(* IEC 61131-3 sources: LASAL/Class/Varan_Base, 1 file *)

(* ---- Varan_Base.st ---- *)
#ifndef _T_VARANBASE_H
#define _T_VARANBASE_H

#define	VARAN_PLL_OFFSET		16#0140
#define VARAN_MULTIPLE_OFFSET	16#01AC

// version of serial number validation (16#10 = 1.0)
#define SERNO_VALIDATION_VERSION 16#10

#define IsTransparent_IS_AVAILABLE

// Defines for Mutex Generation
#define VARAN_STR_MUTEX_NAME_SEPERATOR ".."
#define VARAN_MUTEX_NAME_END_LENGTH 5
#define VARAN_MUTEX_NAME_MAX_LENGTH 32

#define VARAN_SPI_IDENT_LICENCENO_OFFSET    16#14
#define VARAN_SPI_IDENT_HARDWAREVER_OFFSET  16#18

#endif // _T_VARANBASE_H

#include "..\..\Class\HwControl\HwControl.h"
#include "..\..\Source\interfaces\lsl_st_hardwaretree.h"

(*!
<Class
	Name               = "Varan_Base"
	Revision           = "2.15"
	RealtimeTask       = "false"
	CyclicTask         = "false"
	BackgroundTask     = "false"
	Sigmatek           = "true"
	OSInterface        = "false"
	HighPriority       = "false"
	Automatic          = "false"
	UpdateMode         = "Prescan"
	IconPath           = ".\Class\Varan_Base\tool.ICO"
	SharedCommandTable = "true"
	Objectsize         = "(468,120)"
	Comment            = "baseclass of varan slave classes">
	<Channels>
		<Server Name="ConnectCounter" Visualized="true" Initialize="false" WriteProtected="true" Retentive="false" Comment="Connects of Module"/>
		<Server Name="DeviceAddress" Visualized="true" Initialize="false" WriteProtected="true" Retentive="false" Comment="device address of hardware module"/>
		<Server Name="DeviceID" Visualized="true" Initialize="false" WriteProtected="true" Retentive="false" Comment="This server shows the device ID of the hardware module."/>
		<Server Name="DiagControl" Visualized="true" Initialize="false" WriteProtected="false" Retentive="false" Comment="Server to control Diagnose Function of module&#13;&#10;&#13;&#10;Read from Server&#13;&#10;-2..wrong FPGA for Diagnose&#13;&#10;-1..wrong OS for Diagnose&#13;&#10;0..Diagnose Function is deaktivated, not available&#13;&#10;1..Diagnose Function activated (additionally you need #define VARAN_DIAGNOSE)&#13;&#10;&#13;&#10;Write to Server&#13;&#10;0..to deactivate Diagnose&#13;&#10;1..to activate Diagnose&#13;&#10;2..to reset Counter (ConnectCounter, FaultCounter, RXLost, TXLost)"/>
		<Server Name="FaultCounter" Visualized="true" Initialize="false" WriteProtected="true" Retentive="false" Comment="PackageCounter for RXLost and TXLost were invalid"/>
		<Server Name="Online" Visualized="true" Initialize="false" WriteProtected="true" Retentive="false" Comment="is class online or not"/>
		<Server Name="Release" Visualized="true" Initialize="false" WriteProtected="true" Retentive="false" Comment="FPGA - Version"/>
		<Server Name="RetryCounter" Visualized="true" Initialize="false" WriteProtected="false" Retentive="false" Comment="retry counter of varan module"/>
		<Server Name="RXLost" Visualized="true" Initialize="false" WriteProtected="true" Retentive="false" Comment="RX-Packages lost"/>
		<Server Name="SerialNo" Class="String" Visualized="true" Initialize="false" WriteProtected="true" Retentive="false" Comment="use this channel to access the string functions"/>
		<Server Name="State" Visualized="true" Initialize="false" WriteProtected="true" Retentive="false" Comment="This server shows the current status of the hardware class. For more information see: Varan hardware class status."/>
		<Server Name="TXLost" Visualized="true" Initialize="false" WriteProtected="true" Retentive="false" Comment="TX-Packages lost"/>
		<Server Name="ValidateSerNo" Visualized="true" Initialize="false" WriteProtected="false" Retentive="false" Comment="if the validation of the serial number is activated (SerNoValidation = 1)&#13;&#10;the serial number of the actual module can be validated by writing to this server&#13;&#10;&#13;&#10;this server shows also the state of validation:&#13;&#10;-2..validation not acivated&#13;&#10;-1..no module validated on this position&#13;&#10; 0..module is not the validated one&#13;&#10; 1..module is the validated one"/>
		<Server Name="VendorID" Visualized="true" Initialize="false" WriteProtected="true" Retentive="false" Comment="This server contains the vendor ID of the hardware module."/>
		<Client Name="Required" Required="true" Internal="false" Comment="0 = module is not required&#13;&#10;1 = module is required (CPU will crash if module is missing)"/>
		<Client Name="SerialNoStr" Required="true" Internal="true"/>
		<Client Name="SerNoBackup" Required="true" Internal="true"/>
		<Client Name="SerNoValidation" Required="false" Internal="false" Comment="0..serial number of varan client does not matter&#13;&#10;1..serial number of varan client has to be validated, to use the module&#13;&#10;&#13;&#10;validation is done via write(1) to the ValidateSerNo Server"/>
		<Client Name="TimeBase" Required="false" Internal="false" DefValue="0"/>
		<Client Name="TimeBaseOffset" Required="false" Internal="false" DefValue="0"/>
		<Client Name="To_MultiTask" Required="false" Internal="false" Comment="This client is automatically connected to a OS interface class."/>
		<Client Name="To_StdLib" Required="false" Internal="false" Comment="This client is automatically connected to a OS interface class."/>
		<Client Name="Transparent" Required="false" Internal="false" DefValue="0" Comment="If this Client is set to 1 the module is not used for building the VARAN-Tree"/>
		<Client Name="UserAction" Required="false" Internal="false" Comment="optional, connect to server to get Varan states via write method.&#13;&#10;possible input values:&#13;&#10; 0..connect&#13;&#10; 1..disconnect&#13;&#10; 2..required data object error&#13;&#10; 3..not required data object error&#13;&#10; 4..fatal error&#13;&#10; 5..time slice error&#13;&#10; 6..watchdog error&#13;&#10; 7..client irq&#13;&#10; 8..device enable&#13;&#10; 9..device disable&#13;&#10;10..irq task interrupt&#13;&#10;11..reactivation of node which was deactivated by software before&#13;&#10;12..irq for direct access alternating buffer (VMC module)&#13;&#10;13..dias error&#13;&#10;14..cdias error (cdias module required behind a CIV)&#13;&#10;&#13;&#10;&#13;&#10;Possible return values:&#13;&#10;0......ok&#13;&#10;&lt;&gt; 0...Generate VaranError&#13;&#10;"/>
		<Client Name="VaranIn" Required="true" Internal="false" Comment="This class must be connected to a VARAN port or a VaranOut_[x] server."/>
	</Channels>
	<Dependencies>
		<Files>
			<File Path=".\Class\VaranManager_Base\VaranManager_Base.h" Include="false"/>
			<File Path=".\Source\interfaces\lsl_st_pci.h" Include="false"/>
			<File Path=".\Class\HwControl\HwControl.h" Include="true"/>
			<File Path=".\Source\interfaces\lsl_st_hardwaretree.h" Include="true"/>
		</Files>
	</Dependencies>
	<RevDoku>
		<Owner Company="Sigmatek" Author="renste"/>
		<Dokumentation Revision="2.15" Date="16.03.2018" Author="EisMic" Company="Sigmatek" Description="Added support for 2nd VaranManager."/>
		<Dokumentation Revision="2.14" Date="06.03.2018" Author="EisMic" Company="Sigmatek" Description="Attached header files no longer point to the installation directory of LASAL but instead now point to the the source/interfaces folder."/>
		<Dokumentation Revision="2.13" Date="10.01.2018" Author="LanSte" Company="Sigmatek" Description="Added Support for default PostInit phase."/>
		<Dokumentation Revision="2.12" Date="23.01.2018" Author="RamAnd" Company="Sigmatek" Description="Log messages have been standardized for easier maintenance, easier use in any class and to allow spam filtering. Code for the logging functions is now only located in HwControl."/>
		<Dokumentation Revision="2.11" Date="28.08.2017" Author="RamAnd" Company="Sigmatek" Description="The NewInst to get hardware diagnosis information doesn&apos;t set the returncode to SPI_ACCESS_FAILED if an optional entry of the type label is not available."/>
		<Dokumentation Revision="2.10" Date="29.11.2016" Author="PieSte" Company="Sigmatek" Description="Changed &quot;Online&quot; server behavior to set online first if cyclic data is valid."/>
		<Dokumentation Revision="2.9" Date="10.05.2016" Author="RamAnd" Company="Sigmatek" Description="Suppressed warning that would occur with target ARM on compiler version 30 or higher."/>
		<Dokumentation Revision="2.8" Date="17.02.2016" Author="EisMic" Company="Sigmatek" Description="Prescalersettings were not set correctly when Payload is active."/>
		<Dokumentation Revision="2.7" Date="28.08.2015" Author="PieSte" Company="Sigmatek" Description="Added support for up to 6 sync outs (e.g. CTMS031) in methode EnableSyncOut()."/>
		<Dokumentation Revision="2.6" Date="17.03.2015" Author="RamAnd" Company="Sigmatek" Description="Added support for Varan Mux."/>
		<Dokumentation Revision="2.5" Date="24.03.2015" Author="EisMic" Company="Sigmatek" Description="Check pointer p_NodeInfo for validity in method GetRetryTimeout due to access exception error if method Varan_HWDisconnect is called and no hardware was available."/>
		<Dokumentation Revision="2.4" Date="28.08.2014" Author="EisMic" Company="Sigmatek" Description="Don&apos;t set states in GetHWInfoData. CMD_Get_Hardware_Diagnosis: Don&apos;t do a return when one spi access failed, try the other IDs too."/>
		<Dokumentation Revision="2.3" Date="24.06.2014" Author="LanSte" Company="Sigmatek" Description="Added support for reading hardware diagnosis."/>
		<Dokumentation Revision="2.2" Date="05.05.2014" Author="LanSte" Company="Sigmatek" Description="Minimized the interface request via CILGET by useing private pointers to reduce time in init."/>
		<Dokumentation Revision="2.1" Date="14.04.2014" Author="RamAnd" Company="Sigmatek" Description="Added new Interface Varan_HwSubBusReady which is called by OS as soon as it has finished enumerating the connected devices on available subbusses."/>
		<Dokumentation Revision="2.0" Date="04.12.2013" Author="RamAnd&#13;&#10;FucHer&#13;&#10;LanSte" Company="Sigmatek" Description="Removed domain support&#13;&#10;Changed AWL code to Structured Text.&#13;&#10;Added Payload Support&#13;&#10;Added include for PCI accesses, which is necessary to find out if the Varan Manager supports LongDOs."/>
		<Dokumentation Revision="1.90" Date="30.08.2013" Author="RamAnd" Company="Sigmatek" Description="The class could have change the state to _DisableError after the disconnect from VARAN, even if there was no further problem."/>
		<Dokumentation Revision="1.80" Date="01.08.2013" Author="LanSte" Company="Sigmatek" Description="Added Support for changeable Payload DO&apos;s"/>
		<Dokumentation Revision="1.70" Date="18.07.2013" Author="LanSte&#13;&#10;ZoePat" Company="Sigmatek" Description="Added Payload Support&#13;&#10;Check if manager is on at function GetNodeInfo() to get different states for connected and disconnected modules if manager is turned off (e.g.: in case of required error that was handled by client UserAction)"/>
		<Dokumentation Revision="1.60" Date="07.03.2013" Author="RamAnd" Company="Sigmatek" Description="Improved comment of client UserAction (added new reasons)"/>
		<Dokumentation Revision="1.50" Date="05.11.2012" Author="RamAnd&#13;&#10;RamAnd" Company="Sigmatek" Description="Corrected time measurement for internal tests.&#13;&#10;Removed resetting of the FPGA retry counter in method ResetDataObject which could result in a wrong behavior of the RetryCounter server."/>
		<Dokumentation Revision="1.40" Date="18.09.2012" Author="RamAnd" Company="Sigmatek" Description="New State &quot;_NoCalibDataFound&quot; if a pointer to calibration data is fetched and there are no calibration data on the client."/>
		<Dokumentation Revision="1.39" Date="18.07.2012" Author="ObeChr" Company="Sigmatek" Description="Implemented time measurement for internal tests in methods UpdateRt, UpdateRtPostScan and UpdateCy&#13;&#10;Reduction of PCI Accesses in Methode GetRetryTimeout()"/>
		<Dokumentation Revision="1.38" Date="09.12.2011" Author="RamAnd" Company="Sigmatek" Description="The actual domain number is now added to the hardware path."/>
		<Dokumentation Revision="1.37" Date="19.09.2011" Author="RamAnd" Company="Sigmatek" Description="The client UserAction can now also be used to prevent a required error, if the write-method of the connected Server returns 0."/>
		<Dokumentation Revision="1.36" Date="13.07.2011" Author="RamAnd" Company="Sigmatek" Description="Added a dependency to class Hub_Base_Root, otherwise crashes can happen if only single VARAN-classes have been updated."/>
		<Dokumentation Revision="1.35" Date="14.04.2011" Author="BleErn" Company="Sigmatek" Description="Set complex object &quot;SerialNoStr&quot; to visualized"/>
		<Dokumentation Revision="1.34" Date="02.03.2011" Author="RamAnd" Company="Sigmatek" Description="Added new input parameter to method SetMultipleDataPointers to handle more than 1 multiple read write commands per VARAN client."/>
		<Dokumentation Revision="1.33" Date="04.01.2011" Author="BleErn" Company="Sigmatek" Description="Added Client Transparent that allows to disable a VARAN-HW-Class"/>
		<Dokumentation Revision="1.32" Date="17.01.2011" Author="RamAnd" Company="Sigmatek" Description="A required error on the first connect of the device can now be detected via the UserAction client"/>
		<Dokumentation Revision="1.31" Date="11.01.2011" Author="RamAnd" Company="Sigmatek" Description="Error fixed that Diagnostic functions stopped working after the first fault occured."/>
		<Dokumentation Revision="1.30" Date="14.12.2010" Author="RamAnd" Company="Sigmatek" Description="Set all servers to visualized, so that they can be used in visualisation"/>
		<Dokumentation Revision="1.29" Date="02.09.2010" Author="BleErn" Company="Sigmatek" Description="Server SerNoValidation was always set to 0 on disconnect of module"/>
		<Dokumentation Revision="1.28" Date="02.08.2010" Author="RamAnd" Company="Sigmatek" Description="Reworked serial number validation, because of problems with non-Sigmatek devices. Now the serial number is saved as a string instead of a number."/>
		<Dokumentation Revision="1.27" Date="22.07.2010" Author="WocPet / RamAnd" Company="Sigmatek" Description="Added functionality to forward a required error.&#13;&#10;Removed client UseRtPostScan (not needed, since it PostScan is always used)"/>
		<Dokumentation Revision="1.26" Date="06.04.2010" Author="RamAnd" Company="Sigmatek" Description="Added method &quot;FlexInit&quot; to initialize class if the position on VARAN has changed (FlexHub functionality)"/>
		<Dokumentation Revision="1.25" Date="10.03.2010" Author="RamAnd" Company="Sigmatek" Description="Added serial number validation and method CheckDeviceID for easier overloading"/>
		<Dokumentation Revision="1.24" Date="04.03.2010" Author="BleErn" Company="Sigmatek" Description="RtPostScan could be disabled at every CIV (took no notice of define!)"/>
		<Dokumentation Revision="1.23" Date="23.02.2010" Author="BleErn" Company="Sigmatek" Description="Changes in handling of VaranRtPostScan"/>
		<Dokumentation Revision="1.22" Date="17.05.2010" Author="RamAnd" Company="Sigmatek" Description="Changed defines to avoid compiler warning &quot;Identical Redefinition&quot;"/>
		<Dokumentation Revision="1.21" Date="09.10.2009" Author="ObeChr" Company="Sigmatek" Description="Added functions for VaranDiagnose"/>
		<Dokumentation Revision="1.20" Date="02.09.2009" Author="RamAnd" Company="Sigmatek" Description="Added functions for safety and hardwaretree."/>
		<Dokumentation Revision="1.19" Date="05.08.2009" Author="ObeChr" Company="Sigmatek" Description="When Client is required and no VaranInterface is available, VaranManager set application into reset"/>
		<Dokumentation Revision="1.18" Date="20.07.2009" Author="ObeChr" Company="Sigmatek" Description="Added function to set run state of do depending on required"/>
		<Dokumentation Revision="1.17" Date="16.07.2009" Author="ObeChr" Company="Sigmatek" Description="Added funktion to use VaranRtPostScan"/>
		<Dokumentation Revision="1.16" Date="18.06.2009" Author="EbnAnt" Company="Sigmatek" Description="Set Varan_CallBack() to virtual"/>
		<Dokumentation Revision="1.15" Date="16.04.2009" Author="RamAnd" Company="Sigmatek" Description="Added new method GetDocumentation to fetch pdf documentation of client.&#13;&#10;Added new Server SerialNo, to display the serial no of varan clients."/>
		<Dokumentation Revision="1.14" Date="01.12.2008" Author="RamAnd" Company="Sigmatek" Description="added new input variable b_use_divider_sync to function EnableSyncOut.&#13;&#10;Corrected SetNewPllData to new address mapping.&#13;&#10;improved client comments"/>
		<Dokumentation Revision="1.13" Date="03.09.2008" Author="renste" Company="Sigmatek" Description="add function for new pll"/>
	</RevDoku>
	<Network Name="Varan_Base">
		<!-- List of Components in this network -->
		<Components>
			<Object
				Name       = "SerialNoStr"
				Class      = "String"
				Position   = "(180,480)"
				Visualized = "true">
				<Channels>
					<Server Name="Data"/>
					<Client Name="SingleRealloc" Value="1"/>
				</Channels>
			</Object>
			<Object
				Name       = "SerNoBackup"
				Class      = "RamFile"
				Position   = "(180,630)"
				Visualized = "true">
				<Channels>
					<Server Name="FileNameHex"/>
					<Server Name="m_udLength"/>
					<Server Name="SizeError"/>
					<Client Name="Alarm"/>
					<Client Name="MultiTask"/>
					<Client Name="Setup" Value="2#1101"/>
				</Channels>
			</Object>
		</Components>
		<Comments>
		</Comments>
		<!-- List of Connections in this network -->
		<Connections>
			<Connection Source="this.SerialNoStr" Destination="SerialNoStr.Data"/>
			<Connection Source="this.SerialNo" Destination="SerialNoStr.Data" Vertices="(818,570),(496,570),"/>
			<Connection Source="this.SerNoBackup" Destination="SerNoBackup.m_udLength"/>
		</Connections>
		<!-- Headerfiles -->
		<Options>
		</Options>
	</Network>
</Class>
*)
Varan_Base : CLASS
	TYPE
	  t_CallBack : STRUCT
	    ud_Counter : UDINT;
	    ud_ConnectCnt : UDINT;
	    ud_DisconnectCnt : UDINT;
	    ud_InterruptCnt : UDINT;
	    ud_SubBusReadyCnt : UDINT;
	    p_InterruptHandleDO : ^LSL_VARANFRAME;  //! <Type Comment="Warning:&#13;&#10;If the Interface &quot;IMULTIVARANMANAGER&quot; is used (b_PayloadSupport = true) this pointer those not point to the DO in the DPRAM!&#13;&#10;In this case this pointer holds the handle to the DO.&#13;&#10;" Name="t_CallBack.p_InterruptHandleDO"/>
	    ud_LastReason : UDINT;
	  END_STRUCT;
	  t_CycleWork :
	  (
	    _CycleInitIdle,
	    _CycleStartAsyDO,
	    _CycleStartIsoDO,
	    _CycleWaitforValidData,
	    _CyclePreOperational,
	    _CycleOperational
	  )$UDINT;
	  t_PllDataRead : STRUCT
	    us_State : BSINT
	    [
	      1 Pll_Locked,
	      2 Pll_Unlocked,
	      3 SyncOutputAvailable0,
	      4 SyncOutputAvailable1,
	      5 SyncOutputAvailable2,
	      6 IRQWatchdogEnable,
	      7 Pll_Enable,
	      8 PeriodeOverwriteAllowed,
	    ];
	  END_STRUCT;
	  t_PllDO : STRUCT
	    p_Handle : ^LSL_VARANFRAME;
	    p_DOSettings : ^t_VaranDOSettingsRd;
	    p_DataRead : ^t_PllDataRead;
	  END_STRUCT;
#pragma pack(push, 1)
	  t_PllSyncOut : STRUCT
	    sd_Offset : DINT;
	    us_PeriodMultiplier : USINT;
	    us_FrameCountTreshold : USINT;
	    us_Reserved1 : USINT;
	    us_ControlStatus : BSINT
	    [
	      1 SyncOutEnable,
	      2 FrameCountEnable,
	      3 SystemSync,  //! <Type Comment="0..divider sync&#13;&#10;1..system sync" Name="t_PllSyncOut.us_ControlStatus.SystemSync"/>
	    ];
	  END_STRUCT;
#pragma pack(pop)
	  t_RootDependency : ^Hub_Base_Root;
#pragma pack(push, 1)
	  t_SerNoValidateHeader : STRUCT
	    Version : HSINT;  //! <Type Comment="X.Y starting with 1.0 as first valid version&#13;&#10;&#13;&#10;X = Major&#13;&#10;Y = Minor" Name="t_SerNoValidateHeader.Version"/>
	    ZeroByte : USINT;
	    StringLength : UDINT;
	  END_STRUCT;
#pragma pack(pop)
	  t_SPI_CalibHeader : STRUCT
	    ud_Checksum : UDINT;
	    ud_ListVersion : UDINT;
	    ud_ListLength : UDINT;
	  END_STRUCT;
	  t_TempDataRead : STRUCT
	    si_Periode : INT;
	    ui_Prescaler : UINT;
	    ui_HiTimeRegister : UINT;
	  END_STRUCT;
	  t_TransparentInfo : BSINT
	  [
	    1 DeviceIsTransparent,
	    2 ClientTransparentRead,
	  ];
	END_TYPE
  //Servers:
	State 	: SvrChCmd_t_e_VaranErrors;
	Online 	: SvrCh_DINT;
	Release 	: SvrCh_HDINT;
	DeviceAddress 	: SvrCh_HDINT;
	VendorID 	: SvrCh_UDINT;
	DeviceID 	: SvrCh_UDINT;
	SerialNo 	: SvrChCmd_UDINT;
	RetryCounter 	: SvrCh_UDINT;
	ValidateSerNo 	: SvrCh_DINT;
	DiagControl 	: SvrCh_DINT;
	ConnectCounter 	: SvrCh_UDINT;
	FaultCounter 	: SvrCh_UDINT;
	RXLost 	: SvrCh_UDINT;
	TXLost 	: SvrCh_UDINT;
  //Clients:
	VaranIn 	: CltChCmd_Hub_Base;
	Required 	: CltCh_DINT;
	UserAction 	: CltCh_DINT;
	SerNoValidation 	: CltCh_DINT;
	Transparent 	: CltCh_DINT;
	To_StdLib 	: CltChCmd__StdLib;
	To_MultiTask 	: CltChCmd__MultiTask;
	TimeBase 	: CltCh_UDINT;
	TimeBaseOffset 	: CltCh_UDINT;
	SerialNoStr 	: CltChCmd_String;
	SerNoBackup 	: CltChCmd_RamFile;
  //Variables:
		ud_VaranManagerNr 	: UDINT;
		pVaran 	: ^LSL_VARAN;			//! <Variable Comment="Pointer for the Varan interface" Name="pVaran"/>
		pMultiVaran 	: ^LSL_MULTI_VARAN;			//! <Variable Comment="Pointer for the MultiVaran/payload support interface" Name="pMultiVaran"/>
		mt_api 	: ^LSL_MT_TYPE;
		p_VaranPosition 	: ^USINT;
		p_NodeInfo 	: ^LSL_VARANNODEINFO;
		s_NodeInfo 	: LSL_VARANNODEINFO;
		ud_HandleModule 	: UDINT;
		ud_DeviceDelayTime 	: UDINT;
		s_CallBackSettings 	: t_CallBack;			//! <Variable Comment="settings of user callback function" Name="s_CallBackSettings"/>
		e_RequiredFaultState 	: t_e_VaranErrors;
		b_DisableDevice 	: BOOL;
		ud_DisableTime 	: UDINT;
		us_MulticastFilter 	: USINT;
		us_MultipleSequence 	: USINT;
		s_TimeRt 	: t_TimeMeasurementVaran;
		s_TimeRtPostScan 	: t_TimeMeasurementVaran;
		s_TimeCy 	: t_TimeMeasurementVaran;
		b_CyTask 	: BOOL;
		p_ObjectPath 	: ^USINT;
		s_Diagnose 	: t_s_VaranDiagnose;
		szSerNoStr : ARRAY [0..SERNO_STRING_SIZE-1] OF CHAR;

		b_ValidationInProgress 	: BOOL;
		SerNoHeader 	: t_SerNoValidateHeader;
		TransparentInfo 	: t_TransparentInfo;
		ud_ResponseTimeMax 	: UDINT;
		b_PayloadSupport 	: BOOL;			//! <Variable Comment="TRUE When Payload DOs are supporded by the OS Interface." Name="b_PayloadSupport"/>
		b_DMAactive 	: BOOL;			//! <Variable Comment="TRUE When Payload DOs are supporded by the OS Interface and the FPGA has an DMA Controller." Name="b_DMAactive"/>
		ud_OffestSPI 	: UDINT;
		bOnline 	: BOOL;
		eCycleWork 	: t_CycleWork;
		uiBasePostInitHandle 	: UINT;
		bPostInitNeeded 	: BOOL;
		_ParaBaseCy 	: CmdStruct;
		_ResultBaseCy 	: results;
  //Functions:
				//! <Function Comment="-------------------------------------------------------------------------------------------------&#13;&#10;[#ENGLISH]&#13;&#10;=================================================================================================&#13;&#10;Construct of Base class to set class not initialized&#13;&#10;=================================================================================================&#13;&#10;[server] State  :W  :State of class&#13;&#10;" Name="Varan_Base"/>
	FUNCTION Varan_Base
		VAR_OUTPUT
			ret_code 	: ConfStates;
		END_VAR;
				//! <Function Comment="Init for Varan Client" Name="Init"/>
	FUNCTION VIRTUAL GLOBAL Init;
				//! <Function Comment="Cy - Funktion of Varan class ( called bei VaranMaster )" Name="UpdateCy"/>
	FUNCTION VIRTUAL GLOBAL UpdateCy;
				//! <Function Comment="Rt - Funktion of Varan class ( called bei VaranMaster )" Name="UpdateRt"/>
	FUNCTION VIRTUAL GLOBAL UpdateRt;
				//! <Function Comment="Function is called by VaranRtPostScan if used" Name="UpdateRtPostScan"/>
	FUNCTION VIRTUAL GLOBAL UpdateRtPostScan;
				//! <Function Comment="get PDF-File from client, if it is available" Name="GetDocumentation"/>
	FUNCTION VIRTUAL GLOBAL GetDocumentation
		VAR_INPUT
			p_dpne 	: ^CHAR;			//! <Variable Comment="pass string of Drive/Path/Name/Extension (e.g. &quot;C:\mydoc.pdf&quot;)" Name="GetDocumentation.p_dpne"/>
		END_VAR
		VAR_OUTPUT
			sd_retval 	: DINT;			//! <Variable Comment=" 0..success&#13;&#10;-1..invalid parameters&#13;&#10;-2..failed to open file&#13;&#10;-3..os version must be 01.02.018 or higher&#13;&#10;-4..no documentation available on this client&#13;&#10;-5..failed to allocate memory for the file content&#13;&#10;-6..error in reading documentation from client&#13;&#10;-7..writing to file failed" Name="GetDocumentation.sd_retval"/>
		END_VAR;
				//! <Function Comment="Function returns pointer to node string of class" Name="GetPointer2NodeString"/>
	FUNCTION VIRTUAL GLOBAL GetPointer2NodeString
		VAR_OUTPUT
			p_us_node 	: ^USINT;			//! <Variable Comment="pointer to node string" Name="GetPointer2NodeString.p_us_node"/>
		END_VAR;
				//! <Function Comment="Function is called if a varan module is connected&#13;&#10;" Name="Varan_HwConnect"/>
	FUNCTION VIRTUAL GLOBAL Varan_HwConnect
		VAR_INPUT
			ud_data 	: UDINT;			//! <Variable Comment="data of callback function" Name="Varan_HwConnect.ud_data"/>
		END_VAR
		VAR_OUTPUT
			sd_retval 	: DINT;			//! <Variable Comment="return value of OS" Name="Varan_HwConnect.sd_retval"/>
		END_VAR;

	FUNCTION Diagnose;
				//! <Function Comment="[#ENGLISH]&#13;&#10;=================================================================================================&#13;&#10;Function to set Pll settings of hardware module&#13;&#10;=================================================================================================&#13;&#10;[server] State    :W  :state of class&#13;&#10;[members] ud_DeviceDelayTime :W  :delay time of varan client for Pll&#13;&#10;   p_NodeInfo   :W  :pointer to varan client informations&#13;&#10;[locals] ud_data    :W/R :data for direct access&#13;&#10;" Name="SetPllData"/>
	FUNCTION SetPllData
		VAR_INPUT
			ud_delay_time 	: UDINT := 0;
		END_VAR
		VAR_OUTPUT
			sd_retval 	: DINT;
		END_VAR;
				//! <Function Comment="[#ENGLISH]&#13;&#10;=================================================================================================&#13;&#10;Function to get device address, Vendor ID and Device ID of varan module&#13;&#10;=================================================================================================&#13;&#10;[server] State   :W  :state of class&#13;&#10;   Release   :W  :FPGA - Version of varan client&#13;&#10;   DeviceAddress :W  :Device Address of client (from os)&#13;&#10;   VendorID  :W  :Vendor ID of varan client&#13;&#10;   DeviceID  :W  :Device ID of varan client&#13;&#10;[members] p_VaranPosition  :R  :node string of varan module&#13;&#10;   p_NodeInfo   :W  :pointer to varan client informations&#13;&#10;[locals] us_pll_time   :W/R :pll time from VaranMaster&#13;&#10;" Name="GetNodeInfo"/>
	FUNCTION GetNodeInfo
		VAR_OUTPUT
			sd_retval 	: DINT;
		END_VAR;
				//! <Function Comment="[#ENGLISH]&#13;&#10;=================================================================================================&#13;&#10;Callback Function is called from VaranManager&#13;&#10;=================================================================================================&#13;&#10;[server] Release   :W  :FPGA - Version of varan client&#13;&#10;   DeviceAddress :W  :Device Address of client (from os)&#13;&#10;   VendorID  :W  :Vendor ID of varan client&#13;&#10;   DeviceID  :W  :Device ID of varan client&#13;&#10;   State   :W  :state of class&#13;&#10;[client] Required  :R  :is class required for varan or not&#13;&#10;   UserAction  :R  :client for user actions&#13;&#10;[members] s_CallBackSettings  :W  :structure for settings of callback function&#13;&#10;   ud_DeviceDelayTime  :W  :delay time of varan client for Pll&#13;&#10;   e_RequiredFaultState :W  :Fault state of class in _RequiredError State&#13;&#10;" Name="Varan_CallBack"/>
	FUNCTION VIRTUAL Varan_CallBack
		VAR_INPUT
			ud_reason 	: UDINT;			//! <Variable Comment="reason of callback" Name="Varan_CallBack.ud_reason"/>
			ud_data 	: UDINT;
		END_VAR
		VAR_OUTPUT
			sd_retval (EAX) 	: DINT;
		END_VAR;
				//! <Function Comment="Function is called if a varan interrupt occures" Name="Varan_HwInterrupt"/>
	FUNCTION VIRTUAL GLOBAL Varan_HwInterrupt
		VAR_INPUT
			ud_reason 	: UDINT;
			ud_data 	: ^t_CallBackInterrupt;
		END_VAR
		VAR_OUTPUT
			sd_retval 	: DINT;
		END_VAR;
				//! <Function Comment="Function is called if a varan module is disconnected&#13;&#10;" Name="Varan_HwDisconnect"/>
	FUNCTION VIRTUAL GLOBAL Varan_HwDisconnect
		VAR_INPUT
			ud_data 	: UDINT;
		END_VAR
		VAR_OUTPUT
			sd_retval 	: DINT;
		END_VAR;

	FUNCTION VIRTUAL GLOBAL Varan_HwSubBusReady
		VAR_INPUT
			ud_data 	: UDINT;
		END_VAR
		VAR_OUTPUT
			sd_retval 	: DINT;
		END_VAR;
				//! <Function Comment="Function to reset settings of a data object" Name="ResetDataObject"/>
	FUNCTION VIRTUAL GLOBAL ResetDataObject
		VAR_INPUT
			p_handleDO 	: ^LSL_VARANFRAME;
			us_state 	: USINT;			//! <Variable Comment="state of DO (cont run, singl run, stop )" Name="ResetDataObject.us_state"/>
			ud_bytes 	: UDINT;			//! <Variable Comment="number of bytes" Name="ResetDataObject.ud_bytes"/>
		END_VAR;
				//! <Function Comment="=================================================================================================&#13;&#10;---------------------- Additional functions------------------------------------------------------&#13;&#10;=================================================================================================&#13;&#10;[#ENGLISH]&#13;&#10;=================================================================================================&#13;&#10;Function to Start time measurement&#13;&#10;=================================================================================================&#13;&#10;" Name="StartTimeMeasurement"/>
	FUNCTION StartTimeMeasurement
		VAR_INPUT
			usMode (EAX) 	: DINT;
		END_VAR;
				//! <Function Comment="[#ENGLISH]&#13;&#10;=================================================================================================&#13;&#10;Function to Stop time measurement&#13;&#10;=================================================================================================&#13;&#10;" Name="StopTimeMeasurement"/>
	FUNCTION StopTimeMeasurement
		VAR_INPUT
			usMode (EAX) 	: DINT;
		END_VAR;
				//! <Function Comment="Function to set a sync out" Name="GetDeviceAddress"/>
	FUNCTION VIRTUAL GLOBAL GetDeviceAddress
		VAR_OUTPUT
			ud_device_address 	: UDINT;			//! <Variable Comment="Device address of client" Name="GetDeviceAddress.ud_device_address"/>
		END_VAR;
				//! <Function Comment="[#ENGLISH]&#13;&#10;=================================================================================================&#13;&#10;Function to set a sync out&#13;&#10;=================================================================================================&#13;&#10;[server] State    :W  :state of class&#13;&#10;[locals] ud_offset    :W/R :address offset in pll&#13;&#10;   p_pll_output_data  :W/R :settings for pll sync output&#13;&#10;" Name="EnableSyncOut"/>
	FUNCTION EnableSyncOut
		VAR_INPUT
			us_sync_nr 	: USINT;			//! <Variable Comment="enable sync0-4 allowed" Name="EnableSyncOut.us_sync_nr"/>
			sd_offset 	: DINT;			//! <Variable Comment="Offset in 10ns time" Name="EnableSyncOut.sd_offset"/>
			us_period_multiplier 	: USINT;			//! <Variable Comment="periode multiplier" Name="EnableSyncOut.us_period_multiplier"/>
			us_frame_count_treshold 	: USINT;			//! <Variable Comment=" Frame Count Treshold" Name="EnableSyncOut.us_frame_count_treshold"/>
			us_enable_frame_count 	: USINT;			//! <Variable Comment=" enable frame count" Name="EnableSyncOut.us_enable_frame_count"/>
			b_use_divider_sync 	: BOOL := FALSE;
		END_VAR
		VAR_OUTPUT
			sd_retval 	: DINT;
		END_VAR;
				//! <Function Comment="Function to get pointer to node information" Name="GetPointer2NodeInfo"/>
	FUNCTION VIRTUAL GLOBAL GetPointer2NodeInfo
		VAR_OUTPUT
			p_node_info 	: ^LSL_VARANNODEINFO;			//! <Variable Comment="Pointer to Node information" Name="GetPointer2NodeInfo.p_node_info"/>
		END_VAR;
				//! <Function Comment="Function to set state of class" Name="SetState"/>
	FUNCTION VIRTUAL GLOBAL SetState
		VAR_INPUT
			sd_error 	: t_e_VaranErrors;			//! <Variable Comment="type of error" Name="SetState.sd_error"/>
		END_VAR;
				//! <Function Comment="Function to disable device" Name="DisableDevice"/>
	FUNCTION VIRTUAL GLOBAL DisableDevice
		VAR_OUTPUT
			sd_retval 	: DINT;
		END_VAR;
				//! <Function Comment="Function to enable device" Name="EnableDevice"/>
	FUNCTION VIRTUAL GLOBAL EnableDevice
		VAR_OUTPUT
			sd_retval 	: DINT;
		END_VAR;
				//! <Function Comment="Function to set all Data Objects off" Name="SetDOsOff"/>
	FUNCTION VIRTUAL GLOBAL SetDOsOff;
				//! <Function Comment="Function to look if class is disabled" Name="IsDeviceDisabled"/>
	FUNCTION VIRTUAL GLOBAL IsDeviceDisabled
		VAR_OUTPUT
			b_disabled 	: BOOL;			//! <Variable Comment="TRUE -&gt; Device is disabled" Name="IsDeviceDisabled.b_disabled"/>
		END_VAR;
				//! <Function Comment="Function to set multiple memory read/write options" Name="SetMultipleSettings"/>
	FUNCTION VIRTUAL GLOBAL SetMultipleSettings
		VAR_INPUT
			us_filter 	: USINT;			//! <Variable Comment="filter of multicast write" Name="SetMultipleSettings.us_filter"/>
			us_sequence 	: USINT;			//! <Variable Comment="sequence number of device" Name="SetMultipleSettings.us_sequence"/>
		END_VAR
		VAR_OUTPUT
			sd_retval 	: DINT;
		END_VAR;
				//! <Function Comment="Function must be overwrite" Name="SetMultipleDataPointers"/>
	FUNCTION VIRTUAL GLOBAL SetMultipleDataPointers
		VAR_INPUT
			p_handle 	: ^LSL_VARANFRAME;			//! <Variable Comment="pointer to data object header" Name="SetMultipleDataPointers.p_handle"/>
			p_data_read 	: ^UDINT;			//! <Variable Comment="pointer to read data" Name="SetMultipleDataPointers.p_data_read"/>
			p_data_write 	: ^UDINT;			//! <Variable Comment="pointer to data write" Name="SetMultipleDataPointers.p_data_write"/>
			DOIndex 	: UDINT;
		END_VAR
		VAR_OUTPUT
			sd_retval 	: DINT;
		END_VAR;
				//! <Function Comment="[#ENGLISH]&#13;&#10;=================================================================================================&#13;&#10;Function to get pointer to calib data&#13;&#10;=================================================================================================&#13;&#10;" Name="GetCalibDataPointer"/>
	FUNCTION GetCalibDataPointer
		VAR_INPUT
			p_offset 	: ^UDINT;			//! <Variable Comment="pointer to variable to write offset" Name="GetCalibDataPointer.p_offset"/>
		END_VAR
		VAR_OUTPUT
			sd_retval 	: DINT;
		END_VAR;
				//! <Function Comment="[#ENGLISH]&#13;&#10;=================================================================================================&#13;&#10;Function to get pointer to calib data&#13;&#10;=================================================================================================&#13;&#10;" Name="ReadSPIData"/>
	FUNCTION ReadSPIData
		VAR_INPUT
			ud_offset 	: UDINT;			//! <Variable Comment="offset in SPI - Flash" Name="ReadSPIData.ud_offset"/>
			ud_length 	: UDINT;			//! <Variable Comment="length of data" Name="ReadSPIData.ud_length"/>
			p_data 	: ^USINT;			//! <Variable Comment="pointer to allocated data space" Name="ReadSPIData.p_data"/>
		END_VAR
		VAR_OUTPUT
			sd_retval 	: DINT;
		END_VAR;
				//! <Function Comment="Function to update module retry counter" Name="UpdateRetryCounter"/>
	FUNCTION VIRTUAL GLOBAL UpdateRetryCounter;
				//! <Function Comment="Function to get varan time" Name="GetVaranTime"/>
	FUNCTION VIRTUAL GLOBAL GetVaranTime
		VAR_INPUT
			p_ud_IsoStartPoint 	: ^UDINT := NIL;
		END_VAR
		VAR_OUTPUT
			ud_varan_time 	: UDINT;			//! <Variable Comment="varan time" Name="GetVaranTime.ud_varan_time"/>
		END_VAR;
				//! <Function Comment="Function to get retry timeout for a number of bytes" Name="GetRetryTimeout"/>
	FUNCTION VIRTUAL GLOBAL GetRetryTimeout
		VAR_INPUT
			ud_bytes 	: UDINT;
		END_VAR
		VAR_OUTPUT
			ud_timeout 	: UDINT;			//! <Variable Comment="retry timout time" Name="GetRetryTimeout.ud_timeout"/>
		END_VAR;
				//! <Function Comment="[#ENGLISH]&#13;&#10;=================================================================================================&#13;&#10;Function to disable Device in Rt (because VARAN_iSetNodeEnableStatus must not called in Realtime)&#13;&#10;=================================================================================================&#13;&#10;" Name="DisableDeviceRt"/>
	FUNCTION DisableDeviceRt
		VAR_OUTPUT
			sd_retval 	: DINT;
		END_VAR;

	FUNCTION SetNewPllData
		VAR_INPUT
			ud_delay_time 	: UDINT := 0;
			us_divider 	: USINT := 0;
		END_VAR
		VAR_OUTPUT
			sd_retval 	: DINT;
		END_VAR;
				//! <Function Comment="Function to set state depending on required" Name="SetRunStatus"/>
	FUNCTION GLOBAL SetRunStatus
		VAR_INPUT
			state 	: USINT;
		END_VAR
		VAR_OUTPUT
			us_retval 	: USINT;
		END_VAR;

	FUNCTION VIRTUAL GLOBAL GetPointer2ObjectPath
		VAR_OUTPUT
			p_us_ObjectPath 	: ^USINT;
		END_VAR;

	FUNCTION VIRTUAL GLOBAL SetObjectThisp
		VAR_INPUT
			p_us_ObjectPath 	: ^USINT;
			ud_thisp 	: UDINT;
		END_VAR
		VAR_OUTPUT
			sd_retval 	: DINT;
		END_VAR;

	FUNCTION VIRTUAL GLOBAL GetObjectThisp
		VAR_INPUT
			p_us_ObjectPath 	: ^USINT;
		END_VAR
		VAR_OUTPUT
			ud_Thisp 	: UDINT;
		END_VAR;

	FUNCTION SerNoValidationTask;

	FUNCTION GetHWInfoData
		VAR_INPUT
			p_offset 	: ^UDINT;
			ud_id 	: UDINT;
		END_VAR
		VAR_OUTPUT
			sd_retval 	: DINT;
		END_VAR;

	FUNCTION GetPllState
		VAR_OUTPUT
			pllstate 	: BSINT;
		END_VAR;

	FUNCTION VIRTUAL CheckCyclicPostInitFinished
		VAR_INPUT
			bForcePostInitEnd 	: BOOL;
		END_VAR;
				//! <Function Comment="Check if DeviceID is supported by class" Name="CheckDeviceID"/>
	FUNCTION VIRTUAL GLOBAL CheckDeviceID
		VAR_INPUT
			ID2Check 	: UDINT;			//! <Variable Comment="VARAN DeviceID, which should be checked" Name="CheckDeviceID.ID2Check"/>
		END_VAR
		VAR_OUTPUT
			IsOK 	: BOOL;			//! <Variable Comment="TRUE...DeviceID is ok with this class&#13;&#10;FALSE..DeviceID is not ok with this class" Name="CheckDeviceID.IsOK"/>
		END_VAR;

	FUNCTION GLOBAL FlexInit;

	FUNCTION GLOBAL AllowRequiredError;

	FUNCTION GLOBAL IsTransparent
		VAR_OUTPUT
			isTransparent 	: BOOL;
		END_VAR;
				//! <Function Comment="Method to add a read payload data object to varan manager.&#13;&#10;The parameters are passed on to the varan manager via a new inst call.&#13;&#10;" Name="AddRdPayloadDO"/>
	FUNCTION VIRTUAL GLOBAL AddRdPayloadDO
		VAR_INPUT
			ud_dol_type 	: UDINT;			//! <Variable Comment="DOL into witch the DO is to be inserted. &#13;&#10;VARAN_DOL_ASY or VARAN_DOL_ISO" Name="AddRdPayloadDO.ud_dol_type"/>
			p_ud_handle 	: ^UDINT;			//! <Variable Comment="Pointer to variable to set the DO handle.&#13;&#10;Value does not represent a valid address." Name="AddRdPayloadDO.p_ud_handle"/>
			ud_offset_read 	: UDINT;			//! <Variable Comment="Offset of read data within the module. &#13;&#10;(DeviceAddress is not included in this value.)" Name="AddRdPayloadDO.ud_offset_read"/>
			ud_length_read 	: UDINT;			//! <Variable Comment="Length of read data object." Name="AddRdPayloadDO.ud_length_read"/>
			p_ud_data_read 	: ^UDINT;			//! <Variable Comment="The pointer to the read data is written to this address." Name="AddRdPayloadDO.p_ud_data_read"/>
			ud_type 	: UDINT := VM_MEMORY_ACCESS;			//! <Variable Comment="0=control area, 1=memory area" Name="AddRdPayloadDO.ud_type"/>
			ud_priority 	: UDINT := VM_PRIORITY_INVALID;			//! <Variable Comment="Priority of the DO within the DOL. &#13;&#10;1000 highest priority&#13;&#10;9000 lowest priority&#13;&#10;Priority not dividable by 1000 cannot be used outside of the init phase.&#13;&#10;Optional." Name="AddRdPayloadDO.ud_priority"/>
			ud_WritePayloadType 	: UDINT := 0;			//! <Variable Comment="Changeable DO.&#13;&#10;Set this parameter if the DO length and or offset needs to be changed after creation.&#13;&#10;Optional." Name="AddRdPayloadDO.ud_WritePayloadType"/>
		END_VAR
		VAR_OUTPUT
			sd_retval 	: DINT;			//! <Variable Comment="Value &lt;&gt; 0 equal an error.&#13;&#10;See &#13;&#10;lsl_st_varan.h   // Ergebniscodes&#13;&#10;VaranManager_Base.h // Return Codes of the Control NewInst method&#13;&#10;for errorcodes." Name="AddRdPayloadDO.sd_retval"/>
		END_VAR;
				//! <Function Comment="Method to add a write payload data object to varan manager.&#13;&#10;The parameters are passed on to the varan manager via a new inst call.&#13;&#10;" Name="AddWrPayloadDO"/>
	FUNCTION VIRTUAL GLOBAL AddWrPayloadDO
		VAR_INPUT
			ud_dol_type 	: UDINT;			//! <Variable Comment="DOL into witch the DO is to be inserted. &#13;&#10;VARAN_DOL_ASY or VARAN_DOL_ISO" Name="AddWrPayloadDO.ud_dol_type"/>
			p_ud_handle 	: ^UDINT;			//! <Variable Comment="Pointer to variable to set the DO handle.&#13;&#10;Value does not represent a valid address." Name="AddWrPayloadDO.p_ud_handle"/>
			ud_offset_write 	: UDINT;			//! <Variable Comment="Offset of write data within the module. &#13;&#10;(DeviceAddress is not included in this value.)" Name="AddWrPayloadDO.ud_offset_write"/>
			ud_length_write 	: UDINT;			//! <Variable Comment="Length of write data object." Name="AddWrPayloadDO.ud_length_write"/>
			p_ud_data_write 	: ^UDINT;			//! <Variable Comment="The pointer to the read data is written to this address." Name="AddWrPayloadDO.p_ud_data_write"/>
			ud_type 	: UDINT;			//! <Variable Comment="0=control area, 1=memory area" Name="AddWrPayloadDO.ud_type"/>
			ud_priority 	: UDINT := VM_PRIORITY_INVALID;			//! <Variable Comment="Priority of the DO within the DOL. &#13;&#10;1000 highest priority&#13;&#10;9000 lowest priority&#13;&#10;Priority not dividable by 1000 cannot be used outside of the init phase.&#13;&#10;Optional." Name="AddWrPayloadDO.ud_priority"/>
			ud_WritePayloadType 	: UDINT := 0;			//! <Variable Comment="Changeable DO.&#13;&#10;Set this parameter if the DO length and or offset needs to be changed after creation.&#13;&#10;Optional." Name="AddWrPayloadDO.ud_WritePayloadType"/>
		END_VAR
		VAR_OUTPUT
			sd_retval 	: DINT;			//! <Variable Comment="Value &lt;&gt; 0 equal an error.&#13;&#10;See &#13;&#10;lsl_st_varan.h   // Ergebniscodes&#13;&#10;VaranManager_Base.h // Return Codes of the Control NewInst method&#13;&#10;for errorcodes." Name="AddWrPayloadDO.sd_retval"/>
		END_VAR;
				//! <Function Comment="Method to add a read/write payload data object to varan manager.&#13;&#10;The parameters are passed on to the varan manager via a new inst call.&#13;&#10;" Name="AddRdWrPayloadDO"/>
	FUNCTION VIRTUAL GLOBAL AddRdWrPayloadDO
		VAR_INPUT
			ud_dol_type 	: UDINT;			//! <Variable Comment="DOL into witch the DO is to be inserted. &#13;&#10;VARAN_DOL_ASY or VARAN_DOL_ISO" Name="AddRdWrPayloadDO.ud_dol_type"/>
			p_ud_handle 	: ^UDINT;			//! <Variable Comment="Pointer to variable to set the DO handle.&#13;&#10;Value does not represent a valid address." Name="AddRdWrPayloadDO.p_ud_handle"/>
			ud_offset_read 	: UDINT;			//! <Variable Comment="Offset of read data within the module. &#13;&#10;(DeviceAddress is not included in this value.)" Name="AddRdWrPayloadDO.ud_offset_read"/>
			ud_length_read 	: UDINT;			//! <Variable Comment="Length of read data object." Name="AddRdWrPayloadDO.ud_length_read"/>
			p_ud_data_read 	: ^UDINT;			//! <Variable Comment="The pointer to the read data is written to this address." Name="AddRdWrPayloadDO.p_ud_data_read"/>
			ud_offset_write 	: UDINT;			//! <Variable Comment="Offset of write data within the module. &#13;&#10;(DeviceAddress is not included in this value.)" Name="AddRdWrPayloadDO.ud_offset_write"/>
			ud_length_write 	: UDINT;			//! <Variable Comment="Length of write data object." Name="AddRdWrPayloadDO.ud_length_write"/>
			p_ud_data_write 	: ^UDINT;			//! <Variable Comment="The pointer to the read data is written to this address." Name="AddRdWrPayloadDO.p_ud_data_write"/>
			ud_type 	: UDINT;			//! <Variable Comment="0=control area, 1=memory area" Name="AddRdWrPayloadDO.ud_type"/>
			ud_priority 	: UDINT := VM_PRIORITY_INVALID;			//! <Variable Comment="Priority of the DO within the DOL. &#13;&#10;1000 highest priority&#13;&#10;9000 lowest priority&#13;&#10;Priority not dividable by 1000 cannot be used outside of the init phase.&#13;&#10;Optional." Name="AddRdWrPayloadDO.ud_priority"/>
			ud_WritePayloadType 	: UDINT := 0;			//! <Variable Comment="Changeable DO.&#13;&#10;Set this parameter if the DO length and or offset needs to be changed after creation.&#13;&#10;Optional." Name="AddRdWrPayloadDO.ud_WritePayloadType"/>
		END_VAR
		VAR_OUTPUT
			sd_retval 	: DINT;			//! <Variable Comment="Value &lt;&gt; 0 equal an error.&#13;&#10;See &#13;&#10;lsl_st_varan.h   // Ergebniscodes&#13;&#10;VaranManager_Base.h // Return Codes of the Control NewInst method&#13;&#10;for errorcodes." Name="AddRdWrPayloadDO.sd_retval"/>
		END_VAR;
				//! <Function Comment="Method to add a move payload data object to varan manager.&#13;&#10;The parameters are passed on to the varan manager via a new inst call.&#13;&#10;" Name="AddMovePayloadDO"/>
	FUNCTION VIRTUAL GLOBAL AddMovePayloadDO
		VAR_INPUT
			ud_dol_type 	: UDINT;			//! <Variable Comment="DOL into witch the DO is to be inserted. &#13;&#10;VARAN_DOL_ASY or VARAN_DOL_ISO" Name="AddMovePayloadDO.ud_dol_type"/>
			p_ud_handle 	: ^UDINT;			//! <Variable Comment="Pointer to variable to set the DO handle.&#13;&#10;Value does not represent a valid address." Name="AddMovePayloadDO.p_ud_handle"/>
			ud_SourceReadDOHandle 	: UDINT;			//! <Variable Comment="Handle of the source DO.&#13;&#10;" Name="AddMovePayloadDO.ud_SourceReadDOHandle"/>
			ud_SourceReadOffset 	: UDINT := 0;			//! <Variable Comment="Offset within the source DO from where to copy the data.&#13;&#10;This offset + the number of bytes to be copied must not exceed the size of the source DO." Name="AddMovePayloadDO.ud_SourceReadOffset"/>
			ud_DestinationWriteDOHandle 	: UDINT;			//! <Variable Comment="Handle of the destination DO.&#13;&#10;" Name="AddMovePayloadDO.ud_DestinationWriteDOHandle"/>
			ud_DestinationWriteOffset 	: UDINT := 0;			//! <Variable Comment="Offset within the destination DO from where to copy the data.&#13;&#10;This offset + the number of bytes to be copied must not exceed the size of the source DO." Name="AddMovePayloadDO.ud_DestinationWriteOffset"/>
			ud_LengthMove 	: UDINT;			//! <Variable Comment="Number of bytes to be copied." Name="AddMovePayloadDO.ud_LengthMove"/>
			ud_Priority 	: UDINT;			//! <Variable Comment="Priority of the DO within the DOL. &#13;&#10;1000 highest priority&#13;&#10;9000 lowest priority&#13;&#10;Priority not dividable by 1000 cannot be used outside of the init phase.&#13;&#10;This value must be set in correct relation with the source and destination DO." Name="AddMovePayloadDO.ud_Priority"/>
		END_VAR
		VAR_OUTPUT
			sd_retval 	: DINT;			//! <Variable Comment="Value &lt;&gt; 0 equal an error.&#13;&#10;See &#13;&#10;lsl_st_varan.h   // Ergebniscodes&#13;&#10;VaranManager_Base.h // Return Codes of the Control NewInst method&#13;&#10;for errorcodes." Name="AddMovePayloadDO.sd_retval"/>
		END_VAR;
				//! <Function Comment="Starts the passed data object " Name="EnableDO"/>
	FUNCTION VIRTUAL GLOBAL EnableDO
		VAR_INPUT
			ud_DOHandle 	: UDINT;			//! <Variable Comment="Starts the passed data object " Name="EnableDO.ud_DOHandle"/>
			ud_bytes 	: UDINT := 0;
		END_VAR
		VAR_OUTPUT
			sd_retval 	: DINT;
		END_VAR;
				//! <Function Comment="Stops the passed data object " Name="DisableDO"/>
	FUNCTION VIRTUAL GLOBAL DisableDO
		VAR_INPUT
			ud_DOHandle 	: UDINT;
			ud_bytes 	: UDINT := 0;
		END_VAR
		VAR_OUTPUT
			sd_retval 	: DINT;
		END_VAR;
				//! <Function Comment="Returns the retry counter of the passed data object." Name="GetRetryCounter"/>
	FUNCTION VIRTUAL GLOBAL GetRetryCounter
		VAR_INPUT
			ud_DOHandle 	: UDINT;
		END_VAR
		VAR_OUTPUT
			us_RetryCounter 	: USINT;
		END_VAR;
				//! <Function Comment="This method is used to change the offset and length of the DO. The method can only be used with the Interface &quot;IMULTIVARANMANAGER&quot; is active (if b_payload). Do not set parameters that are unused/should remain unchanged." Name="ChangeDOLengthOffset"/>
	FUNCTION VIRTUAL GLOBAL ChangeDOLengthOffset
		VAR_INPUT
			ud_DOHandle 	: UDINT;			//! <Variable Comment="Handle of the DO" Name="ChangeDOLengthOffset.ud_DOHandle"/>
			ud_offset_read 	: UDINT := VM_DO_PROPERTY_INVALID;			//! <Variable Comment="New read offset" Name="ChangeDOLengthOffset.ud_offset_read"/>
			ud_length_read 	: UDINT := VM_DO_PROPERTY_INVALID;			//! <Variable Comment="New read length" Name="ChangeDOLengthOffset.ud_length_read"/>
			ud_offset_write 	: UDINT := VM_DO_PROPERTY_INVALID;			//! <Variable Comment="New write offset" Name="ChangeDOLengthOffset.ud_offset_write"/>
			ud_length_write 	: UDINT := VM_DO_PROPERTY_INVALID;			//! <Variable Comment="New write length" Name="ChangeDOLengthOffset.ud_length_write"/>
		END_VAR
		VAR_OUTPUT
			sd_retval 	: DINT;
		END_VAR;

	FUNCTION VIRTUAL GLOBAL SetPrescaler
		VAR_INPUT
			ud_DOHandle 	: UDINT;
			Prescaler 	: UDINT;
			PrescalerCnt 	: UDINT := 0;
			b_MultipleTimeBase 	: BOOL := false;
		END_VAR
		VAR_OUTPUT
			sd_retval 	: DINT;
		END_VAR;
				//! <Function Comment="Install callback function&#13;&#10;&#13;&#10;Overload the method if the derived class needs its own Callback Method. See VDM085, VDM086 for example." Name="InstallCallbackObject"/>
	FUNCTION VIRTUAL InstallCallbackObject
		VAR_OUTPUT
			sd_retval 	: DINT;
		END_VAR;

	FUNCTION VIRTUAL GLOBAL CreateMutex
		VAR_INPUT
			MutexName 	: ^CHAR;
			pThis 	: ^VirtualBase := nil;
		END_VAR
		VAR_OUTPUT
			pv_RetMutex 	: pVoid;
		END_VAR;

	FUNCTION VIRTUAL GLOBAL MutexStart
		VAR_INPUT
			pMutex 	: pVoid;
		END_VAR;

	FUNCTION VIRTUAL GLOBAL MutexStop
		VAR_INPUT
			pMutex 	: pVoid;
		END_VAR;
				//! <Function Comment="Method simulates a SingleRun DO by En/Disabling the DO depending on p_b_DOIsRunning.&#13;&#10;To use this method t_SingleRunState^.StartRequest must be set where the singlerun is required&#13;&#10;and the Method must be called at the end of the task where the DO is used. (UpdatyCy, UpdateRt...)&#13;&#10;Only works with Varan DO (No with Mover)&#13;&#10;Method was made for Payload DO. Should work with standard DO&apos;s as well.&#13;&#10;(EnableDO, DisableDO does not equal ResetDO!)" Name="SingleRunSM"/>
	FUNCTION VIRTUAL GLOBAL SingleRunSM
		VAR_INPUT
			p_DOhandle 	: ^UDINT;
			p_b_DOIsRunning 	: ^t_SingleRunState;
		END_VAR;

	FUNCTION VIRTUAL GLOBAL ChangeMovDOLengthOffset
		VAR_INPUT
			ud_MovDOHandle 	: UDINT;
			ud_SourceReadDOHandle 	: UDINT := VM_DO_PROPERTY_INVALID;
			ud_SourceReadOffset 	: UDINT := VM_DO_PROPERTY_INVALID;
			ud_DestinationWriteDOHandle 	: UDINT := VM_DO_PROPERTY_INVALID;
			ud_DestinationWriteOffset 	: UDINT := VM_DO_PROPERTY_INVALID;
			ud_LengthMove 	: UDINT := VM_DO_PROPERTY_INVALID;
		END_VAR
		VAR_OUTPUT
			sd_retval 	: DINT;
		END_VAR;

	FUNCTION VIRTUAL GLOBAL GetDeviceID
		VAR_OUTPUT
			output 	: UDINT;
		END_VAR;

	FUNCTION VIRTUAL GetFWVersion
		VAR_INPUT
			pData 	: ^CHAR;
			length 	: UDINT;
		END_VAR;
				//! <Function Comment="Returns true if this class needs the postinitphase. &#13;&#10;Default in the base is false." Name="CheckPostInitNeeded"/>
	FUNCTION VIRTUAL GLOBAL CheckPostInitNeeded
		VAR_INPUT
			pbPostInitSettings 	: ^t_VM_CMD_NEED_POST_INIT_CALL_SETTINGS;
		END_VAR
		VAR_OUTPUT
			PostInitNeeded 	: BOOL;
		END_VAR;

	FUNCTION VIRTUAL LogError
		VAR_INPUT
			e_msg 	: ^CHAR;
		END_VAR;

	FUNCTION VIRTUAL LogValue
		VAR_INPUT
			pString 	: ^CHAR;
			Value 	: UDINT;
			Value2 	: UDINT := 16#FFFFFFFF;
			Value3 	: UDINT := 16#FFFFFFFF;
		END_VAR;

	FUNCTION VIRTUAL GLOBAL State::NewInst
		VAR_INPUT
			pPara 	: ^CmdStruct;
			pResult 	: ^results;
		END_VAR
		VAR_OUTPUT
			ret_code 	: iprStates;
		END_VAR;

	FUNCTION VIRTUAL GLOBAL ValidateSerNo::Write
		VAR_INPUT
			input (EAX) 	: DINT;
		END_VAR
		VAR_OUTPUT
			result (EAX) 	: DINT;
		END_VAR;

	FUNCTION VIRTUAL GLOBAL DiagControl::Write
		VAR_INPUT
			input (EAX) 	: DINT;
		END_VAR
		VAR_OUTPUT
			result (EAX) 	: DINT;
		END_VAR;
  //Tables:
	FUNCTION @STD
		VAR_OUTPUT
			ret_code	: CONFSTATES;
		END_VAR;
	FUNCTION GLOBAL TAB @CT_;
END_CLASS;

#pragma using RamFile
#pragma using String
#pragma usingLtd _MultiTask
#pragma usingLtd _StdLib
#pragma usingLtd Hub_Base

#pragma usingLtd Hub_Base_Root

(************************************************************************************
*
*	Baseclass for varan mastercontrolling
*	Created : Sigmatek	/	SR	/	March-April 2006
*	Changes :
*
*
*     FOR NEWER CHANGES SEE REVISION DOCUMENTATION IN CLASS PROPERTIES
*
*   1.11 => 1.12	/	26.05.2008
*			- [DB 863]: - add function to disable device in cyclic
*       1.10 => 1.11 /  18.04.2008
*			- [DB 852]: extend method GetVaranTime to get the IsoStartPoint
*		1.9 => 1.10	/	04.12.2007
*			- [DB 561]:	only call Init of this class (not virtual init)
*		1.8 => 1.9	/	18.07.2007
*			- [DB 561]:	Add function to read Varan time
*			- [DB 632]:	Ignore Execute Fault of Admin - Task with Disable - Function
*			- [DB 594]: set methode GetRetryTimout to global
*		1.7 => 1.8	/	11.07.2007
*			- [DB 620]:	Insert function to update module retry counters
*		1.6 => 1.7	/ 	04.04.2007
*			- [DB 541]: insert function to read SPI data
*			- [DB 536]: interrogation if Fault Boot - Image of FPGA is active
*		1.5 => 1.6	/	13.03.2007
*			- [DB 526]:	only search for position string if no string pointer is available
*		1.4 => 1.5	/	05.02.2007
*			- [DB 493]: changes in function GetDeviceAddress (do not request class state)
*			- Set DisableDevice Flag back if RTOS - Version <= 1.1.141
*		1.3 => 1.4	/	29.01.2007
*			- [DB 461]: add multiple read/write command
*		1.2 => 1.3	/	03.01.2007
*			- [DB 418]: insert functions to disable and enable port
*		1.1 => 1.2	/	14.12.2006
*			- [DB 441]: add function to set state of class
*		1.0 => 1.1	/	28.11.2006
*			first library version
*		0.2 => 1.0	/	05.10.2006
*			initial version
*		0.1 => 0.2	/	13.06.2006
*			second testversion
*		0.0	=> 0.1	/	10.04.2006
*			first testversion for fair in Hannover
*
************************************************************************************)

VAR_PRIVATE

  // Private pointers to interface to avoid multiple OS_CILGet calls.
  pMultiVaranFetch : ^LSL_MULTI_VARAN;
  mt_apiFetch      : ^LSL_MT_TYPE;

  p_this            : ^void;

  //Private Variables for CMD_GET_HARDWARE_DIAGNOSIS AND CMD_GET_HARDWARE_TREE_ENTRY
  a_HWTEntryStr     : ARRAY[0.. VARAN_MAX_DEPTH+1] OF CHAR;  // VaranMaxDepth +1 because length is 2 byte long
  a_VendorName			: ARRAY[0..99] OF CHAR;
  a_DeviceName			: ARRAY[0..99] OF CHAR;
  a_OrderingNoId	  : ARRAY[0..99] OF CHAR;
  a_IdentList_LicenseNo_HwRev   : ARRAY[0..99] OF CHAR;
  a_FWVersion           : ARRAY[0..99] OF CHAR;
  a_SerialNo			: ARRAY[0..31] OF CHAR;

END_VAR

//[#ENGLISH]
//=================================================================================================
//Construct of Base class to set class not initialized
//=================================================================================================
//[server]	State		:W		:State of class
FUNCTION  Varan_Base::Varan_Base
  VAR_OUTPUT
    ret_code		: CONFSTATES;
  END_VAR

  State			:= _NotInitialized;
  ret_code		:= C_OK;

#ifdef HWC_LogInit
  HWC_LogInit();
#endif

  pMultiVaranFetch := nil;
  mt_apiFetch := nil;

END_FUNCTION //  Varan_Base::Varan_Base
//[#ENGLISH]
//=================================================================================================
//Init for Varan Client
//=================================================================================================
//[server]	State				:W		:state of class
//[client]	Required			:R		:is class required for varan or not
//[members]	p_VaranPosition		:R/W	:node string of varan module
//			ud_VaranManagerNr	:W		:number of varan manager
//			p_Varan				:W		:pointer to varan OS - Functions
//[locals]	sd_retval			:W/R	:return value of called functions
FUNCTION VIRTUAL GLOBAL Varan_Base::Init
  VAR
    sd_retval	: DINT;
#ifdef VARAN_DIAGNOSE
    dummy     : UDINT;
#endif
    // For NewInst command
    _Para 	            : CmdStruct;
    _Result 	          : Results;
    ret_code            : IprStates;
    paraGetModuleHandel : t_VM_CMD_GetModuleHandle;
    b_DummyCallback     : BOOL;
    bPostInitSettings   : t_VM_CMD_NEED_POST_INIT_CALL_SETTINGS;
  END_VAR

//=================================================================================================
#ifdef VM_CLASS_TIME_MEASUREMENT
    s_TimeRt.ud_MaximalTime := 0;
    s_TimeRt.ud_MinimalTime := 16#FFFF_FFFF;

    s_TimeRtPostScan.ud_MaximalTime := 0;
    s_TimeRtPostScan.ud_MinimalTime := 16#FFFF_FFFF;

    s_TimeCy.ud_MaximalTime := 0;
    s_TimeCy.ud_MinimalTime := 16#FFFF_FFFF;
#endif
//=================================================================================================

  b_DummyCallback := false;

  //read required client
  Required := Required.read() and 1;

  //-----------------------------------------------------------------------------------------------
  // Check if Payload is supported by the VM

  _Para.uiCmd := VM_CMD_SET_MUX_THIS;
  _Para.aPara[0] := this$DINT;

  VaranIn.NewInst(#_Para, #_Result);

  //-----------------------------------------------------------------------------------------------
  // Check if Payload is supported by the VM
  _Para.uiCmd := VM_CMD_IS_PAYLOAD_SUPPORTED;
  _Result.aData[0]$BOOL := 0;   // Set to 0 in case the NewInst Method is not Implemented

  if VaranIn.NewInst(#_Para, #_Result) = READY then
    b_PayloadSupport := _Result.aData[0]$BOOL;
  end_if;

  // Check if the FPGA has (and uses) an DMA Controller
  if b_PayloadSupport then
    _Para.uiCmd := VM_CMD_IS_DMA_ACTIVE;
    _Result.aData[0]$BOOL := 0;   // Set to 0 in case the NewInst Method is not Implemented

    if VaranIn.NewInst(#_Para, #_Result) = READY then
      b_DMAactive := _Result.aData[0]$BOOL;
    end_if;
  end_if;

  //-----------------------------------------------------------------------------------------------
  //get master number
  ud_VaranManagerNr := VaranIn.GetManagerNumber( p_varan := #pVaran );

  //look for an error
  if ( pVaran = NIL ) &
     ( b_PayloadSupport = false ) then  // pVaran is only used without PayloadSupport
    State := _NoVaranInterface;
    if Required then
      VaranIn.AllowRequiredError();
    end_if;
    return;
  end_if;

  //-----------------------------------------------------------------------------------------------
  //get Varan position if we have no position yet
  if ( p_VaranPosition = NIL ) then

    //alloc memory to get position
    p_VaranPosition := ( To_StdLib.Malloc( size := VARAN_MAX_DEPTH + 1 ) )$^USINT;

    //look if an error occurs
    if ( p_VaranPosition = NIL ) then
      State := _RootError;
      return;
    end_if;

    //set length to 0
    p_VaranPosition^ := 0;

    //get position
    sd_retval := VaranIn.GetVaranPosition( p_us_info := p_VaranPosition );

    //look if an error occurs
    if ( sd_retval <> VARANMANAGER_OK ) then
      State := _RootError;

      // if it's connected via flex hub, install a dummy callback before leaving the method
      if (VaranIn.Read() = VM_FLEXHUB_READ_ID) then
        //-----------------------------------------------------------------------------------------------
        //install callback function
        sd_retval := VaranIn.SetObjectCallback	( p_us_position_info	:= NIL
                            , ud_action_ptr			:= ( #Varan_CallBack() )$UDINT
                            , ud_thisp				:= this$UDINT
                            , sd_required			:= Required
                            );

        //look if an error occurs
        if ( sd_retval <> VARANMANAGER_OK ) then
          return;
        else
          // State := _NoHardware;
          State := _NotInitialized; // State to _NotInitialized, Otherwise the derived class will not create the DOs and abort the init.
          b_DummyCallback := true;
        end_if;
      else
        return;
      end_if;
    end_if;

    //alloc memory for position pointer
    p_VaranPosition := 	( To_StdLib.ReAlloc	( mptr		:= p_VaranPosition
                        , newsize	:= p_VaranPosition^ + 1
                        )
              )$^USINT;

    //look if an error occurs
    if ( p_VaranPosition = NIL ) then
      State := _RootError;
      return;
    end_if;

    // Get Module Handle if supported
    if b_PayloadSupport then

      if pMultiVaranFetch = nil then

        // Get the pointer for the Payload inteface
        if ( OS_CILGet( INTERFACE_MULTIVARANMANAGER, #pMultiVaranFetch ) <> SYS_ERR_NONE) then
          // Should be impossible b_PayloadSupport is only set when this interface was already called succesfully
          LogError("@017C (Varan_Base::Init) No Multi_Varan Interface found");
          State 		:= _NoVaranInterface;
          return;
        end_if;

      end_if;

      pMultiVaran := pMultiVaranFetch;

      // Only read Module handle if it has not been read yet
      // May already be read be other classes with the same position string. (For example CDIAS behind CIV)
      if ud_HandleModule = 0 then

        _Para.uiCmd := VM_CMD_GET_MODULE_HANDLE;

        paraGetModuleHandel.p_us_position_info := p_VaranPosition;
        paraGetModuleHandel.p_ud_module_handle := #ud_HandleModule;

        _Para.aPara[0]  := (#paraGetModuleHandel)$DINT;

        if VaranIn.NewInst(#_Para, #_Result) = READY then
          if _result.aData[0]$DINT <> VM_CMD_OK then
            State := _RootError;
            return;
          end_if;
        else
          State := _RootError;
          return;
        end_if;
      end_if;

    end_if;

    // Post Init Support --------------------------------------------------------------------------

    bPostInitSettings := 0; // Init with 0 incase derived classes forget to set parameter.
    bPostInitNeeded   := CheckPostInitNeeded(#bPostInitSettings);
    if bPostInitNeeded then

      _Para.uiCmd     := VM_CMD_NEED_POST_INIT_CALL;
      _Para.aPara[0]  := this$DINT;
      _Para.aPara[1]  := bPostInitSettings$DINT;

      ret_code        := VaranIn.NewInst(pPara:= #_Para, pResult:= #_Result);

      if ret_code = READY then
        uiBasePostInitHandle := _Result.aData[0];
      else
        // PostInit Flag zuruecksetzen da nicht von VM unterstuetzt.
        bPostInitNeeded := FALSE;
        // Keine Trace ausgabe, wird schon im VM gemacht
      end_if;
    end_if;

  end_if;

  //-----------------------------------------------------------------------------------------------
  if b_DummyCallback = false then  // Only install if there is not dummy callback due to not connected module to Flexhub

    //install callback function
    sd_retval := InstallCallbackObject();

    //look if an error occurs
    if ( sd_retval <> VARANMANAGER_OK ) then
      State := _CallBackError;
      return;
    end_if;

  end_if;

  //Get Object Path
  GetPointer2ObjectPath();

#ifdef VARAN_DIAGNOSE
  s_Diagnose.TimeCounter := 1000000 / VaranIn.GetVaranTime(p_ud_IsoStartPoint := #dummy); //value, when we increment every cycle after 1 sec
#endif

END_FUNCTION //VIRTUAL GLOBAL Varan_Base::Init
//[#ENGLISH]
//=================================================================================================
//Rt - Funktion of Varan class ( called bei VaranMaster )
//=================================================================================================
FUNCTION VIRTUAL GLOBAL Varan_Base::UpdateRt

  //disable Device if an error interrupt occures (not in interrupt because it takes to long)
  //if we have a Cy - Task disable Device in cylcic otherwise call special function (VaranManager disables Device in cyclic)
  //if DisableDevice is called in Rt a Timeslice Error can occure because OS uses ADMIN Task for this function!!!
  if (b_CyTask = FALSE) then

    if ( b_DisableDevice = TRUE) then
      DisableDeviceRt();
      SetDOsOff();
    end_if;

    // Check if Cylic Post Init needs to be finished
    if bPostInitNeeded then
      CheckCyclicPostInitFinished(FALSE);
    end_if;

  end_if;

END_FUNCTION //VIRTUAL GLOBAL Varan_Base::UpdateRt
//[#ENGLISH]
//=================================================================================================
//Cy - Funktion of Varan class ( called bei VaranMaster )
//=================================================================================================
FUNCTION VIRTUAL GLOBAL Varan_Base::UpdateCy

  b_CyTask := TRUE;

#ifdef VARAN_DIAGNOSE
  if (s_Diagnose.Command <> Deactivate) & (s_Diagnose.Counter >= s_Diagnose.TimeCounter) & (DiagControl >= 0) then
    Diagnose();
    s_Diagnose.Counter  := 0;
  elsif (s_Diagnose.Command = Deactivate) then
    DiagControl         := 0;
    s_Diagnose.Counter  := 0;
  elsif (DiagControl >= 0) then
    s_Diagnose.Counter    += 1;
  end_if;
#endif

  //disable Device if an error interrupt occures (not in interrupt because it takes to long)
  if ( b_DisableDevice = TRUE ) then
    DisableDevice();
    SetDOsOff();
  end_if;

  // Check if Cylic Post Init needs to be finished
  if bPostInitNeeded then
    CheckCyclicPostInitFinished(FALSE);
  end_if;

END_FUNCTION //VIRTUAL GLOBAL Varan_Base::UpdataCy
//[#ENGLISH]
//=================================================================================================
//Function returns pointer to node string of class
//=================================================================================================
//[members]	p_VaranPosition		:R		:Node string of varan module
//[<p_us_node]pointer to node string
FUNCTION VIRTUAL GLOBAL Varan_Base::GetPointer2NodeString
  VAR_OUTPUT
    p_us_node		: ^USINT;
  END_VAR

  if IsTransparent() then
    p_us_node := NIL; //We have no Nodestring: we do not exist!
  else

    //get Varan position if we have no position yet
    if ( p_VaranPosition = NIL ) then
      Varan_Base::Init();
    end_if;

    p_us_node := p_VaranPosition;

  end_if;

END_FUNCTION //VIRTUAL GLOBAL Varan_Base::GetPointer2NodeString
//[#ENGLISH]
//=================================================================================================
//Function is called if a varan interrupt occures
//=================================================================================================
//[server]	Online					:W		:set if class is ok and all data is valid
//			State					:W		:state of class
//[members]	s_CallBackSettings		:W		:structure for settings of callback function
//[>ud_reason]reason of interrupt
//[>ud_data]data of call back
//[<sd_retval]returnvalue of function
FUNCTION VIRTUAL GLOBAL Varan_Base::Varan_HwInterrupt
  VAR_INPUT
    ud_reason	: UDINT;
    ud_data		: ^t_CallBackInterrupt;
  END_VAR
  VAR_OUTPUT
    sd_retval	: DINT;
  END_VAR

  Online	:= 0;
  bOnline := FALSE;

  //look which type of interrupt
  case ( ud_reason ) of
    VARANMANAGER_CB_REQ_ERROR:
      State			:= _HardwareRequiredIRQ;

    VARANMANAGER_CB_NOT_REQ_ERROR:
      State			:= _HardwareNotRequiredIRQ;
      b_DisableDevice := TRUE;

    VARANMANAGER_FATAL_ERROR:
      State			:= _HardwareFatalErrorIRQ;
      b_DisableDevice	:= TRUE;

  end_case;

  //get pointer to data object with error
  s_CallBackSettings.p_InterruptHandleDO := ( ud_data^.ud_Handle )$^LSL_VARANFRAME;

  sd_retval := VARANMANAGER_OK;

END_FUNCTION //VIRTUAL GLOBAL Varan_Base::Varan_HwInterrupt
//[#ENGLISH]
//=================================================================================================
//Function is called if a varan module is connected
//=================================================================================================
//[server]	Online		:W		:set if class is ok and all data is valid
//			State		:W		:state of class
//[>ud_data]data of call back
//[<sd_retval]returnvalue of function
#pragma warning(disable: 73)

FUNCTION VIRTUAL GLOBAL Varan_Base::Varan_HwConnect
  VAR_INPUT
    ud_data		: UDINT;
  END_VAR
  VAR_OUTPUT
    sd_retval	: DINT;
  END_VAR

  //set Online 1 first if cyclic data is valid
  Online    := 1;
  bOnline   := TRUE;
  State     := _ClassOk;
  sd_retval := VARANMANAGER_OK;

END_FUNCTION //VIRTUAL GLOBAL Varan_Base::Varan_HwConnect
//[#ENGLISH]
//=================================================================================================
//Function is called if a varan module is disconnected
//=================================================================================================
//[server]	Online		:W		:set if class is ok and all data is valid
//			State		:W		:state of class
//[>ud_data]data of call back
//[<sd_retval]returnvalue of function
FUNCTION VIRTUAL GLOBAL Varan_Base::Varan_HwDisconnect
  VAR_INPUT
    ud_data		: UDINT;
  END_VAR
  VAR_OUTPUT
    sd_retval	: DINT;
  END_VAR

  Online		:= 0;
  bOnline   := FALSE;
  State     := _NoHardware;

  if bPostInitNeeded then

    CheckCyclicPostInitFinished(bForcePostInitEnd:=TRUE);

  end_if;

  sd_retval := VARANMANAGER_OK;

END_FUNCTION //VIRTUAL GLOBAL Varan_Base::Varan_HwDisconnect
#pragma warning(default: 73)

//[#ENGLISH]
//=================================================================================================
//Callback Function is called from VaranManager
//=================================================================================================
//[server]	Release			:W		:FPGA - Version of varan client
//			DeviceAddress	:W		:Device Address of client (from os)
//			VendorID		:W		:Vendor ID of varan client
//			DeviceID		:W		:Device ID of varan client
//			State			:W		:state of class
//[client]	Required		:R		:is class required for varan or not
//			UserAction		:R		:client for user actions
//[members] s_CallBackSettings		:W		:structure for settings of callback function
//			ud_DeviceDelayTime		:W		:delay time of varan client for Pll
//			e_RequiredFaultState	:W		:Fault state of class in _RequiredError State
//[<sd_retval]0=Ok, VARANMANAGER_CALLBACK_NOT_HANDLED=VaranError
//[>ud_reason]reason of callback
//[>ud_data]data of callback function
FUNCTION VIRTUAL Varan_Base::Varan_CallBack
  VAR_INPUT
    ud_reason 	: UDINT;
    ud_data 	: UDINT;
  END_VAR
  VAR_OUTPUT
    sd_retval (EAX) 	: DINT;
  END_VAR

  //counter to count number of callback calls
  s_CallBackSettings.ud_Counter += 1;
  s_CallBackSettings.ud_LastReason := ud_reason;

  //switch case of callback
  case ( ud_reason ) of
//**********************************************************************************************************************************************************
    // Interrupt
    VARANMANAGER_CB_REQ_ERROR,
    VARANMANAGER_CB_NOT_REQ_ERROR,
    VARANMANAGER_FATAL_ERROR:
                    sd_retval := Varan_HwInterrupt	( ud_reason := ud_reason
                                                    , ud_data := ud_data$^t_CallBackInterrupt
                                                    );

                    s_CallBackSettings.ud_InterruptCnt += 1;

//**********************************************************************************************************************************************************
    // Connnect of a device
    VARANMANAGER_CB_CONNECT:
                    sd_retval := Varan_HwConnect( ud_data := ud_data );
                    s_CallBackSettings.ud_ConnectCnt += 1;

#ifdef VARAN_DIAGNOSE
                    //Varan Diangose
                    //Init Struct
                    s_Diagnose.cmd_Input.ManagerNr       := ud_VaranManagerNr;               //number of manager
                    s_Diagnose.cmd_Input.BaseAddress     := DeviceAddress;                   //base-address of node
                    s_Diagnose.cmd_Input.CounterLength   := 20;                              //5 counter a 4 byte
                    s_Diagnose.cmd_Input.Counter1        := 0;                               //flags
                    s_Diagnose.cmd_Input.Counter2        := 1;                               //connect_count
                    s_Diagnose.cmd_Input.Counter3        := 2;                               //fault_count
                    s_Diagnose.cmd_Input.Counter4        := 3;                               //rx_lost
                    s_Diagnose.cmd_Input.Counter5        := 4;                               //tx_lost
                    s_Diagnose.InputSize                 := sizeof(s_Diagnose.cmd_Input); //size of input-struct

                    if s_Diagnose.ActiveMerker = TRUE then
                      s_Diagnose.Command := Activate;
                    end_if;

#endif

//**********************************************************************************************************************************************************
    // Disconnect of a device
    VARANMANAGER_CB_DISCONNECT:		sd_retval := Varan_HwDisconnect( ud_data := ud_data );
                    s_CallBackSettings.ud_DisconnectCnt += 1;
                    Release := 0;
                    DeviceAddress := 0;
                    VendorID := 0;
                    DeviceID := 0;
                    ud_DeviceDelayTime := 0;
                    IF ValidateSerNo <> -2 THEN
                      ValidateSerNo := 0;
                    END_IF;
                    SerialNoStr.Clear();

#ifdef VARAN_DIAGNOSE
                    if s_Diagnose.Command = Activate then
                      s_Diagnose.ActiveMerker := TRUE;
                    else
                      s_Diagnose.ActiveMerker := FALSE;
                    end_if;

                    s_Diagnose.Command := Deactivate;
#endif

//**********************************************************************************************************************************************************
    VARANMANAGER_CB_SUB_BUSES_INITIALIZED:
                    sd_retval := Varan_HwSubBusReady( ud_data := ud_data );
                    s_CallBackSettings.ud_SubBusReadyCnt += 1;

//**********************************************************************************************************************************************************
  end_case;

  //------------------------------------------------------------------------------------------------
  //if class is required and state is error (because of first connect (called in Init))
  if 	( Required
    & (State 	<> _ClassOk)
    & (State	<> _NotInitialized)
    & (State	<> _InvalidSerialNo)
    & (State	<> _ModuleFoundButManagerIsOff)
    )
  then

    //give an error back to VaranManager to shut down application
    sd_retval := VARANMANAGER_CALLBACK_NOT_HANDLED;
    //save fault state
    e_RequiredFaultState := State;
    //Set state of class
    State := _RequiredError;

    //Set VaranMaster off
    VaranIn.SetManagerOff( e_error := State );

  else
    //if we have a negative return code but class is not required then we do nothing
    if ( sd_retval <> VARANMANAGER_OK ) then
      sd_retval := VARANMANAGER_OK;
    end_if;
  end_if;

  //----------------------------------User has last word -------------------------------------------
  //look if user client is connected
  if ( IsClientConnected( #UserAction ) = TRUE ) then

    //call user call back so that user has chance to change return value to VaranManager
    if (State = _RequiredError) & (sd_retval = VARANMANAGER_CALLBACK_NOT_HANDLED) then
      sd_retval := UserAction.write( VARANMANAGER_CB_REQ_ERROR );
    else
      sd_retval := UserAction.write( ud_reason$DINT );
    end_if;

    //look if user want other reaction
    if ( sd_retval ) then
      sd_retval := VARANMANAGER_CALLBACK_NOT_HANDLED;
    else
      sd_retval := VARANMANAGER_OK;
    end_if;
  end_if;

END_FUNCTION // Varan_Base::Varan_CallBack
//[#ENGLISH]
//=================================================================================================
//Function to get device address, Vendor ID and Device ID of varan module
//=================================================================================================
//[server]	State			:W		:state of class
//			Release			:W		:FPGA - Version of varan client
//			DeviceAddress	:W		:Device Address of client (from os)
//			VendorID		:W		:Vendor ID of varan client
//			DeviceID		:W		:Device ID of varan client
//[members]	p_VaranPosition		:R		:node string of varan module
//			p_NodeInfo			:W		:pointer to varan client informations
//[locals]	us_pll_time			:W/R	:pll time from VaranMaster
//[<sd_retval]0=OK, else varan manager error
FUNCTION Varan_Base::GetNodeInfo
  VAR_OUTPUT
    sd_retval	: DINT;
  END_VAR
  VAR
    szValidSerNo : ARRAY [0..SERNO_STRING_SIZE-1] OF CHAR;
    ManagerState  : t_e_VaranErrors;
  END_VAR

  if b_PayloadSupport then
    p_NodeInfo := #s_NodeInfo;  // No direct access with payload support, data will be stored to the passed pointer
  end_if;

  //get node info from os
  sd_retval := VaranIn.GetNodeInfo( p_us_position_info	:= p_VaranPosition
                                  , p_node_info			:= #p_NodeInfo
                                  );

  //look for an error
  if ( sd_retval <> VARANMANAGER_OK ) then
    State := _NoHardware;
    return;
  end_if;

  //set class servers
  Release			:= TO_UDINT( p_NodeInfo^.ucFPGAVersion );

  //check for Fault Boot Image version of FPGA
  if ( Release < 16#10 ) then
    State := _ErrorBootImageFPGA;
    sd_retval := -100;
    return;
  end_if;

  DeviceAddress	:= p_NodeInfo^.uiAddress;
  VendorID		:= p_NodeInfo^.uiVendorID;
  DeviceID		:= p_NodeInfo^.uiDeviceID;

  // check device ID before we continue with serial number check
  if CheckDeviceID(DeviceID) = FALSE then
    State := _WrongHardware;
    sd_retval := -101;
    return;
  end_if;

  // check if manager is on
  ManagerState := VaranIn.GetManagerState();
  if ManagerState <> _ClassOk then
    State := _ModuleFoundButManagerIsOff;
    sd_retval := -105;
    return;
  end_if;

  // get serial number of this client (from spi flash)
  VaranIn.GetSerialNo(p_us_position_info:=p_VaranPosition, p_SerialNo:=#szSerNoStr[0]);

  SerialNoStr.WriteDataOff(udLen:=_StrLen(#szSerNoStr[0]), udOff:=0, pData:=#szSerNoStr[0]);

  SerNoValidation := SerNoValidation.Read();
  if SerNoValidation then

    // get header out of ramfile
    if SerNoBackup.GetDataAt(p_us_data:=(#SerNoHeader)$^USINT, ud_size:=sizeof(SerNoHeader), ud_at:=0) = C_OK then

      // initialize local string
      _memset(#szValidSerNo[0], 0, SERNO_STRING_SIZE);

      // check data in header (string must be smaller than string size: 1 byte for termination) and get string out of ramfile
      if (SerNoHeader.Version = 16#10) & (SerNoHeader.ZeroByte = 0) & (SerNoHeader.StringLength < SERNO_STRING_SIZE) &
         (SerNoBackup.GetDataAt(p_us_data:=(#szValidSerNo[0])$^USINT, ud_size:=SerNoHeader.StringLength, ud_at:=sizeof(SerNoHeader)) = C_OK) then

        // check if it's the correct serial number string
        if _strcmp(#szSerNoStr[0], #szValidSerNo[0]) = 0 then
        ValidateSerNo := 1;
      else
          // strings doesn't match
        ValidateSerNo := 0;
        State := _InvalidSerialNo;

          // return errorcode to prevent initialisation of the device
          sd_retval := -104;
      end_if;
    else
      ValidateSerNo := -1;
      State := _InvalidSerialNo;

        // header invalid or failed to read serno string
        sd_retval := -103;
      end_if;
    else
      ValidateSerNo := -1;
      State := _InvalidSerialNo;

      // failed to read header of serno data
      sd_retval := -102;
    end_if;

  else
    ValidateSerNo := -2;
  end_if;

END_FUNCTION //VIRTUAL GLOBAL Varan_Base::GetNodeInfo
//[#ENGLISH]
//=================================================================================================
//Function to reset settings of a data object
//=================================================================================================
//[client]	Required		:R		:is class required for varan or not
//[>p_HandleDO]pointer to data object
//[>us_state]state of DO (cont run, singl run, stop )
//[>ud_bytes]number of bytes in DO
FUNCTION VIRTUAL GLOBAL Varan_Base::ResetDataObject
  VAR_INPUT
    p_handleDO		: ^LSL_VARANFRAME;
    us_state		: USINT;
    ud_bytes		: UDINT;
  END_VAR

  //look if we have a valid pointer
  if ( p_handleDO <> NIL ) then

    //set state of DO
    if ( Required ) then
      p_handleDO^.ucCtrlStat 		:= us_state or VARAN_DO_REQUIRED;
    else
      p_handleDO^.ucCtrlStat 		:= us_state;
    end_if;

    //reset retry counter
//		p_handleDO^.ucRetryCounter	:= 0;

    //set number of allowed retries
    p_handleDO^.ucRetrys		:= VM_ALLOWED_RETRIES;

    //set time for retry timeout
    p_handleDO^.uiRetryTimeout	:= GetRetryTimeout( ud_bytes := ud_bytes );
  end_if;

END_FUNCTION // Varan_Base::ResetDataObject

//[#ENGLISH]
//=================================================================================================
//Function to set Pll settings of hardware module
//=================================================================================================
//[server]	State				:W		:state of class
//[members]	ud_DeviceDelayTime	:W		:delay time of varan client for Pll
//			p_NodeInfo			:W		:pointer to varan client informations
//[locals]	ud_data				:W/R	:data for direct access
//[<sd_retval]0=OK, else varan manager error
FUNCTION Varan_Base::SetPllData
  VAR_INPUT
    ud_delay_time 	: UDINT;
  END_VAR
  VAR_OUTPUT
    sd_retval 	: DINT;
  END_VAR
  VAR
    ud_data			    : UDINT;
  END_VAR

  //calculate right register value (Response Time (in 10ns steps) / 2 - constant FPGA delay time
  ud_DeviceDelayTime := ( p_NodeInfo^.uiResponseTime ) / 20 + VM_CONST_FPGA_DELAY + ud_delay_time;

  //set device delay time and max. value of missing pll input sync
  ud_data := ( ud_DeviceDelayTime shl 8 ) or VM_MAX_PLL_SYNC_MISS;

  // Payload Support
  if b_PayloadSupport then
    //write Pll time with direct access
    sd_retval := MULTI_VARAN_iExecuteDirectAccess(  hNodeHandle := ud_HandleModule
                                                  , udCommand   := VARAN_CMD_CONTROL_WRITE
                                                  , udOffset    := VARAN_PLL_OFFSET + 16#B
                                                  , udLength    := sizeof(ud_data)
                                                  , pusData     := ( #ud_data )$^USINT
                                                  , pudErrorInfo:= NIL);
  else
    //write Pll time with direct access
    sd_retval := VARAN_iWriteControlDA( uiManager		  := ud_VaranManagerNr
                                      , uiAddress		  := DeviceAddress + VARAN_PLL_OFFSET + 16#B
                                      , uiLen			    := sizeof(ud_data)
                                      , uiRetryTimeout:= GetRetryTimeout( ud_bytes := sizeof(ud_data) )
                                      , pvData		    := ( #ud_data )$^UDINT
                                      , puiError		  := NIL
                                      );
  end_if;

  //look if an error occurs
  if ( sd_retval <> VARANMANAGER_OK ) then
    State := _PllError;
    return;
  end_if;

END_FUNCTION //VIRTUAL GLOBAL Varan_Base::SetPllData
//[#ENGLISH]
//=================================================================================================
//Function to set a sync out
//=================================================================================================
//[server]	State				:W		:state of class
//[locals]	ud_offset				:W/R	:address offset in pll
//			p_pll_output_data		:W/R	:settings for pll sync output
//[>us_sync_nr]enable sync0-4 allowed
//[>sd_offset]Offset in 10ns time
//[>us_period_multiplier]periode multiplier
//[>us_frame_count_treshold] Frame Count Treshold
//[>us_enable_frame_count] enable frame count
//[<sd_retval]returnvalue of os
FUNCTION Varan_Base::EnableSyncOut
  VAR_INPUT
    us_sync_nr 	: USINT;
    sd_offset 	: DINT;
    us_period_multiplier 	: USINT;
    us_frame_count_treshold 	: USINT;
    us_enable_frame_count 	: USINT;
    b_use_divider_sync 	: BOOL;
  END_VAR
  VAR_OUTPUT
    sd_retval 	: DINT;
  END_VAR
  VAR
    ud_offset				: UDINT;
    p_pll_output_data		: t_PllSyncOut;
  END_VAR

  //look which sync out we have
  if ( us_sync_nr <= 5 ) then

    ud_offset := 16#10 + ( us_sync_nr * 16#8 );

    //set out data
    p_pll_output_data.sd_Offset 			:= sd_offset;
    p_pll_output_data.us_PeriodMultiplier	:= us_period_multiplier;
    p_pll_output_data.us_FrameCountTreshold	:= us_frame_count_treshold;
    p_pll_output_data.us_Reserved1			:= 0;

    p_pll_output_data.us_ControlStatus.SyncOutEnable 	:= TRUE;
    p_pll_output_data.us_ControlStatus.FrameCountEnable	:= us_enable_frame_count$BOOL;
    p_pll_output_data.us_ControlStatus.SystemSync       := NOT b_use_divider_sync;

    // Payload Support
    if b_PayloadSupport then
      //write Pll time with direct access
      sd_retval := MULTI_VARAN_iExecuteDirectAccess(  hNodeHandle := ud_HandleModule
                                                    , udCommand   := VARAN_CMD_CONTROL_WRITE
                                                    , udOffset    := VARAN_PLL_OFFSET + ud_offset
                                                    , udLength    := sizeof(t_PllSyncOut)
                                                    , pusData     := ( #p_pll_output_data )$^USINT
                                                    , pudErrorInfo:= NIL);
    else
      //write Pll time with direct access
      sd_retval := VARAN_iWriteControlDA	( uiManager		  := ud_VaranManagerNr
                                          , uiAddress		  := DeviceAddress + VARAN_PLL_OFFSET + ud_offset
                                          , uiLen			    := sizeof(t_PllSyncOut)
                                          , uiRetryTimeout:= GetRetryTimeout( ud_bytes := sizeof(t_PllSyncOut) )
                                          , pvData		    := ( #p_pll_output_data )$^UDINT
                                          , puiError		  := NIL
                                          );
    end_if;

    //look if an error occurs
    if ( sd_retval <> VARANMANAGER_OK ) then
      State := _PllError;
      return;
    end_if;

  else
    sd_retval := -100;
  end_if;

END_FUNCTION // Varan_Base::EnableSyncOut
//[#ENGLISH]
//=================================================================================================
//Function to set a sync out
//=================================================================================================
//[server]	DeviceAddress	:W		:Device Address of varan client
//[locals]	sd_retval		:W/R	:return value of called dfunctions
//[<ud_device_address]Device address of client
FUNCTION VIRTUAL GLOBAL Varan_Base::GetDeviceAddress
  VAR_OUTPUT
    ud_device_address	: UDINT;
  END_VAR
  VAR
    sd_retval			: DINT;
  END_VAR

  //look if we have a device address
  if ( DeviceAddress = 0 ) then

    //get node information
    sd_retval := GetNodeInfo();

    //look for an error
    if ( sd_retval <> VARANMANAGER_OK ) then
      return;
    end_if;
  end_if;

  //return Device Address of varan client
  ud_device_address := DeviceAddress;

END_FUNCTION //VIRTUAL GLOBAL Varan_Base::GetDeviceAddress
//[#ENGLISH]
//=================================================================================================
//Function to get pointer to node information
//=================================================================================================
//[members]	p_node_info	:R/W		:pointer to node information of client (from os)
//[locals]	sd_retval	:W/R		:retunr value of called functions
//[<p_node_info]Pointer to Node information
FUNCTION VIRTUAL GLOBAL Varan_Base::GetPointer2NodeInfo
  VAR_OUTPUT
    p_node_info		: ^LSL_VARANNODEINFO;
  END_VAR
  VAR
    sd_retval	: DINT;
  END_VAR

  //look if we have a correct pointer (we must call init and GetNodeInfo - Function)
  if ( p_NodeInfo = NIL ) then

    //if required error do nothing
    if ( State = _RequiredError ) then
      p_node_info := NIL;
      return;
    end_if;

    //call init function
    Varan_Base::Init();

    //get node info
    sd_retval := GetNodeInfo();

    //look for an error
    if ( sd_retval <> VARANMANAGER_OK ) then
      p_node_info := NIL;
      return;
    end_if;
  end_if;

  //return pointer
  p_node_info := p_NodeInfo;

END_FUNCTION //VIRTUAL GLOBAL Varan_Base::GetPointer2NodeInfo
//[#ENGLISH]
//=================================================================================================
//Function to get retry timeout for a number of bytes
//=================================================================================================
//[members]	p_NodeInfo		:R		:pointer to node information of client (from os)
//[>ud_bytes]number of bytes
//[<ud_timeout]retry timout time
FUNCTION GLOBAL Varan_Base::GetRetryTimeout
  VAR_INPUT
    ud_bytes		: UDINT;
  END_VAR
  VAR_OUTPUT
    ud_timeout		: UDINT;
  END_VAR

  //Got already ResponseTime?
  if ud_ResponseTimeMax = 0 then
    if p_NodeInfo then
      ud_ResponseTimeMax := p_NodeInfo^.uiResponseTimeMax;
    end_if;
  end_if;

  ud_timeout := ud_ResponseTimeMax + ud_bytes * VM_TIMEOUT_ONE_BYTE + VM_RETRY_TIMEOUT_STD_OFFSET;

END_FUNCTION // Varan_Base::GetRetryTimeout
//=================================================================================================
//---------------------- Additional functions------------------------------------------------------
//=================================================================================================

//[#ENGLISH]
//=================================================================================================
//Function to Start time measurement
//=================================================================================================
#pragma warning(disable:74)
#pragma warning(disable:73)
FUNCTION Varan_Base::StartTimeMeasurement
  VAR_INPUT
    usMode (EAX) 	: DINT;
  END_VAR
#ifdef VM_CLASS_TIME_MEASUREMENT
  VAR
    tmpTime : ^t_TimeMeasurementVaran;
  END_VAR

  case usMode of

    //-----------------------------------------------------------

    VARANTIME_RT:
      tmpTime := #s_TimeRt;

    //-----------------------------------------------------------

    VARANTIME_RTPOSTSCAN:
      tmpTime := #s_TimeRtPostScan;

    //-----------------------------------------------------------

    VARANTIME_CY:
      tmpTime := #s_TimeCy;

    //-----------------------------------------------------------

  end_case;

  if ( tmpTime^.us_Activate ) then
//    Save_Flg();
    CLI();
    tmpTime^.ud_Timemark := VaranIn.GetNsTime();
  end_if;

#endif

END_FUNCTION // Varan_Base::StartTimeMeasurement
//[#ENGLISH]
//=================================================================================================
//Function to Stop time measurement
//=================================================================================================
FUNCTION Varan_Base::StopTimeMeasurement
  VAR_INPUT
    usMode (EAX) 	: DINT;
  END_VAR
#ifdef VM_CLASS_TIME_MEASUREMENT
  VAR
    tmpTime : ^t_TimeMeasurementVaran;
  END_VAR

  case usMode of

    //-----------------------------------------------------------

    VARANTIME_RT:
      tmpTime := #s_TimeRt;

    //-----------------------------------------------------------

    VARANTIME_RTPOSTSCAN:
      tmpTime := #s_TimeRtPostScan;

    //-----------------------------------------------------------

    VARANTIME_CY:
      tmpTime := #s_TimeCy;

    //-----------------------------------------------------------

  end_case;

  if ( tmpTime^.us_Activate ) then

    //get actual time
    tmpTime^.ud_ActualTime := VaranIn.GetNsTime() - tmpTime^.ud_Timemark;

    //look for maximum time
    if ( tmpTime^.ud_ActualTime > tmpTime^.ud_MaximalTime ) then
      tmpTime^.ud_MaximalTime := tmpTime^.ud_ActualTime;
    end_if;

    //look for minimum time
    if ( tmpTime^.ud_ActualTime < tmpTime^.ud_MinimalTime ) then
      tmpTime^.ud_MinimalTime := tmpTime^.ud_ActualTime;
    end_if;

    //look for average time (100000 cycles)
    if ( tmpTime^.ud_AverageCounter = 100000 ) then

      tmpTime^.ud_AverageTime 	:= tmpTime^.ud_AverageSum / tmpTime^.ud_AverageCounter;
      tmpTime^.ud_AverageSum 	:= 0;
      tmpTime^.ud_AverageCounter := 0;

    else
      tmpTime^.ud_AverageSum += ( tmpTime^.ud_ActualTime / 100 );
      tmpTime^.ud_AverageCounter += 1;
    end_if;

    STI();
//    Restore_Flg();
  end_if;

#endif

END_FUNCTION // Varan_Base::StopTimeMeasurement
#pragma warning(default:74)
#pragma warning(default:73)

//[#ENGLISH]
//=================================================================================================
//Function to set state of class
//=================================================================================================
//[>sd_error]type of error
FUNCTION VIRTUAL GLOBAL Varan_Base::SetState
  VAR_INPUT
    sd_error		: t_e_VaranErrors;
  END_VAR

  //only set error if class is ok
  if ( State = _ClassOk ) then

    State := sd_error;

  else
    //only eeprom error can be cleared
    if ( State = _EEPromError & sd_error = _ClassOk ) then
      State := sd_error;
    end_if;
  end_if;

END_FUNCTION //VIRTUAL GLOBAL Varan_Base::SetState
//[#ENGLISH]
//=================================================================================================
//Function to disable device
//=================================================================================================
//[<sd_retval]0=ok, -17=Port no link, -30=client disabled, -31=client cant enable, -100 function not available with this os version, other return code of os
FUNCTION VIRTUAL GLOBAL Varan_Base::DisableDevice
  VAR_OUTPUT
    sd_retval	: DINT;
  END_VAR
  VAR
    nodeProperty    : LSL_PROPERTY_VALUE_PAIR;
  END_VAR

  //look if funtion is available with this os version
  if ( _RTOSVersion >= VM_DISABLE_DEVICE_AVAILABLE ) then

    if b_PayloadSupport then
      nodeProperty.udPropertyId    := ND_PROP_CONNECTION_STATE;
      nodeProperty.udPropertyValue := CN_STATE_DISCONNECTED;
      sd_retval := MULTI_VARAN_iSetNodeProperties(  hNodeHandle           := ud_HandleModule
                                                  , udPropertyCount       := 1
                                                  , psPropertyValuePairs  := #nodeProperty);
    else
      //disable device
      sd_retval := VARAN_iSetNodeEnableStatus	( uiManager		:= ud_VaranManagerNr
                          , pucNode		:= p_VaranPosition
                          , uiNodeStatus	:= 0
                          );
    end_if;

    // if there was an error at disabling it was not caused by a disabled previous module
    if	( sd_retval <> VARANMANAGER_OK ) &
        ( sd_retval <> VARANMANAGER_CLIENT_DISABLED ) &
        ( sd_retval <> VARANMANAGER_ADMIN_DOL_EXECUTION_ERROR	) &	//because if device before is disabled, DA can't work
        ( VaranIn.IsDeviceDisabled() = FALSE ) then

      State := _DisableError;

      //Set VaranMaster off
      VaranIn.SetManagerOff( e_error := State );
    end_if;

    //port is disabled
    b_DisableDevice := FALSE;
    ud_DisableTime := ops.tAbsolute;
  else
    b_DisableDevice := FALSE;
    sd_retval := -100;
  end_if;
